(* IEC 61131-3 sources: plc_NativeGateway/tests, 8 files *)

(* ---- NG_TimeResponseTest.st ---- *)
FUNCTION_BLOCK NG_TimeResponseTest
VAR_OUTPUT
    Done : BOOL;
    Passed : UINT;
    FailedChecks : UINT;
    CaseCount : UINT;
END_VAR
VAR
    Parser : NG_JsonParse;
    Reader : NG_TimeResponse;
    Doc : NG_Document;
    Bytes : NG_Bytes;
    CopyString : STRING_TO_BUF;
    Payload : STRING[2048];
    Stage : UINT;
    CaseIndex : UINT := 1;
    Expected : BOOL;
    Retained : BOOL;
    Actual : BOOL;
END_VAR
IF Done THEN RETURN; END_IF;
Parser(Execute:=Stage=1,Length:=TO_UDINT(LEN(Payload)),Buffer:=Bytes,Doc:=Doc);
CASE Stage OF
0:
    CASE CaseIndex OF
        1: Payload:='{"schemaVersion":1,"gatewayId":"PLC-01","requestId":"time-boot-A-1","bootId":"boot-A","sessionId":"session-A","clientMonoMs":10000,"serverReceivedAt":1792739100000,"serverSentAt":1792739100005}'; Expected:=TRUE; Retained:=FALSE;
        2: Payload:='{"schemaVersion":1,"gatewayId":"PLC-01","requestId":"time-boot-A-1","bootId":"boot-A","sessionId":"session-A","clientMonoMs":10000,"serverReceivedAt":1792739100000,"serverSentAt":1792739100005}'; Expected:=TRUE; Retained:=FALSE;
        3: Payload:='{"schemaVersion":1,"gatewayId":"PLC-01","requestId":"time-boot-A-1","bootId":"boot-A","sessionId":"session-A","clientMonoMs":10000,"timestamp":0,"serverReceivedAt":1792739100000,"serverSentAt":1792739100005}'; Expected:=FALSE; Retained:=FALSE;
        4: Payload:='{"schemaVersion":1,"gatewayId":"PLC-01","requestId":"time-boot-A-1","bootId":"boot-A","sessionId":"session-A","clientMonoMs":true,"serverReceivedAt":1792739100000,"serverSentAt":1792739100005}'; Expected:=FALSE; Retained:=FALSE;
        5: Payload:='{"schemaVersion":1,"gatewayId":"PLC-01","requestId":"time-boot-A-1","bootId":"boot-A","sessionId":"session-A","clientMonoMs":10000.0,"serverReceivedAt":1792739100000,"serverSentAt":1792739100005}'; Expected:=FALSE; Retained:=FALSE;
        6: Payload:='{"schemaVersion":1.0,"gatewayId":"PLC-01","requestId":"time-boot-A-1","bootId":"boot-A","sessionId":"session-A","clientMonoMs":10000,"serverReceivedAt":1792739100000,"serverSentAt":1792739100005}'; Expected:=FALSE; Retained:=FALSE;
        7: Payload:='{"schemaVersion":1,"gatewayId":"PLC-01","requestId":"time-boot-A-1","bootId":"boot-A","sessionId":null,"clientMonoMs":10000,"serverReceivedAt":1792739100000,"serverSentAt":1792739100005}'; Expected:=FALSE; Retained:=FALSE;
        8: Payload:='{"schemaVersion":1,"gatewayId":"PLC-01","requestId":"time-boot-A-1","bootId":"boot-A","sessionId":"session-A","clientMonoMs":9007199254740992,"serverReceivedAt":1792739100000,"serverSentAt":1792739100005}'; Expected:=FALSE; Retained:=FALSE;
        9: Payload:='{"schemaVersion":1,"gatewayId":"PLC-01","requestId":"aaaaaaaaaaaaaaaaaaaaaaaaaaaaaaaaaaaaaaaaaaaaaaaaaaaaaaaaaaaaaaaaa","bootId":"boot-A","sessionId":"session-A","clientMonoMs":10000,"serverReceivedAt":1792739100000,"serverSentAt":1792739100005}'; Expected:=FALSE; Retained:=FALSE;
        10: Payload:='{"schemaVersion":1,"gatewayId":"PLC-01","requestId":"a/b","bootId":"boot-A","sessionId":"session-A","clientMonoMs":10000,"serverReceivedAt":1792739100000,"serverSentAt":1792739100005}'; Expected:=FALSE; Retained:=FALSE;
        11: Payload:='{"schemaVersion":1,"gatewayId":"PLC-01","requestId":"time-boot-A-1","bootId":"boot-A","sessionId":"session-A","clientMonoMs":10000,"serverReceivedAt":1792739100000,"serverSentAt":1792739100005}'; Expected:=FALSE; Retained:=TRUE;
        12: Payload:='{"schemaVersion":1,"gatewayId":"other","requestId":"time-boot-A-1","bootId":"boot-A","sessionId":"session-A","clientMonoMs":10000,"serverReceivedAt":1792739100000,"serverSentAt":1792739100005}'; Expected:=FALSE; Retained:=FALSE;
        13: Payload:='{"schemaVersion":1,"gatewayId":"PLC-01","requestId":"time-boot-A-1","bootId":"other","sessionId":"session-A","clientMonoMs":10000,"serverReceivedAt":1792739100000,"serverSentAt":1792739100005}'; Expected:=FALSE; Retained:=FALSE;
        14: Payload:='{"schemaVersion":1,"gatewayId":"PLC-01","requestId":"time-boot-A-1","bootId":"boot-A","sessionId":"other","clientMonoMs":10000,"serverReceivedAt":1792739100000,"serverSentAt":1792739100005}'; Expected:=FALSE; Retained:=FALSE;
        15: Payload:='{"schemaVersion":1,"gatewayId":"PLC-01","requestId":"other","bootId":"boot-A","sessionId":"session-A","clientMonoMs":10000,"serverReceivedAt":1792739100000,"serverSentAt":1792739100005}'; Expected:=FALSE; Retained:=FALSE;
        16: Payload:='{"schemaVersion":1,"gatewayId":"PLC-01","requestId":"time-boot-A-1","bootId":"boot-A","sessionId":"session-A","clientMonoMs":10001,"serverReceivedAt":1792739100000,"serverSentAt":1792739100005}'; Expected:=FALSE; Retained:=FALSE;
        17: Payload:='{"schemaVersion":1,"gatewayId":"PLC-01","requestId":"time-boot-A-1","bootId":"boot-A","sessionId":"session-A","clientMonoMs":10000.0,"serverReceivedAt":1792739100000,"serverSentAt":1792739100005}'; Expected:=FALSE; Retained:=FALSE;
        18: Payload:='{"schemaVersion":1,"gatewayId":"PLC-01","requestId":"time-boot-A-1","bootId":"boot-A","sessionId":"session-A","clientMonoMs":10000,"serverReceivedAt":1792739100000,"serverSentAt":1.0}'; Expected:=FALSE; Retained:=FALSE;
        19: Payload:='{"schemaVersion":1,"gatewayId":"PLC-01","requestId":"time-boot-A-1","bootId":"boot-A","sessionId":"session-A","clientMonoMs":10000,"serverReceivedAt":1792739100000,"serverSentAt":9007199254740992}'; Expected:=FALSE; Retained:=FALSE;
        20: Payload:='{"schemaVersion":1,"gatewayId":"PLC-01","requestId":"time-boot-A-1","bootId":"boot-A","sessionId":"session-A","clientMonoMs":10000,"serverReceivedAt":true,"serverSentAt":1792739100005}'; Expected:=FALSE; Retained:=FALSE;
        21: Payload:='{"schemaVersion":1,"gatewayId":"PLC-01","requestId":"time-boot-A-1","bootId":"boot-A","sessionId":"session-A","clientMonoMs":10000,"serverReceivedAt":1792739100000,"serverSentAt":1792739100005,"timestamp":0}'; Expected:=FALSE; Retained:=FALSE;
        22: Payload:='{"schemaVersion":1,"gatewayId":"PLC-01","requestId":"time-boot-A-1","bootId":"boot-A","sessionId":"session-A","clientMonoMs":10000,"serverReceivedAt":1792739100000,"serverSentAt":1792739100005,"schemaVersion":1}'; Expected:=FALSE; Retained:=FALSE;
        23: Payload:='{"schemaVersion":1e0,"gatewayId":"PLC-01","requestId":"time-boot-A-1","bootId":"boot-A","sessionId":"session-A","clientMonoMs":10000,"serverReceivedAt":1792739100000,"serverSentAt":1792739100005}'; Expected:=FALSE; Retained:=FALSE;
    END_CASE;
    CopyString(REQ:=FALSE,BUF_FORMAT:=FALSE,BUF_OFFS:=0,BUF_CNT:=LEN(Payload),SRC:=Payload,BUFFER:=Bytes);
    CopyString(REQ:=TRUE,BUF_FORMAT:=FALSE,BUF_OFFS:=0,BUF_CNT:=LEN(Payload),SRC:=Payload,BUFFER:=Bytes);
    IF CopyString.DONE THEN Stage:=1; END_IF;
1:
    IF Parser.Error OR Parser.Done THEN
        Actual:=FALSE;
        IF Parser.Done THEN
            Reader(Length:=TO_UDINT(LEN(Payload)),Retained:=Retained,GatewayId:='PLC-01',BootId:='boot-A',
                SessionId:='session-A',RequestId:='time-boot-A-1',ClientMonoMs:=10000,Doc:=Doc,Bytes:=Bytes);
            Actual:=Reader.Valid;
        END_IF;
        IF Actual=Expected THEN Passed:=Passed+1; ELSE FailedChecks:=FailedChecks+1; END_IF;
        CaseCount:=CaseCount+1; Stage:=2;
    END_IF;
2:
    CaseIndex:=CaseIndex+1;
    IF CaseIndex>23 THEN Done:=TRUE; ELSE Stage:=0; END_IF;
END_CASE;
END_FUNCTION_BLOCK

(* ---- audit_facts_test.st ---- *)
PROGRAM Main
VAR
    Buffer : NG_Buffer;
    Event : NG_CaptureEvent;
    AuditRecord : NG_AuditEvent;
    Cursor : NG_SourceCursor;
    Capture : NG_CaptureCore;
    Poll : NG_PollSlot;
    Audit : NG_AuditCapture;
    Decide : NG_AuditDecision;
    Policy : NG_ReportPolicy;
    Checks : ARRAY[1..20] OF BOOL;
    Passed : UINT;
    FailedChecks : UINT;
    Done : BOOL;
    i : UINT;
END_VAR
(* Compile-only harness; no socket, SDK, persistent store, RTC or physical I/O.
   Cold compilation does not execute these assertions. *)
IF Done THEN RETURN; END_IF;
Checks[1]:=SIZEOF(Event)=UDINT#72;
Checks[2]:=SIZEOF(AuditRecord)=UDINT#80;
Checks[3]:=SIZEOF(Cursor)=UDINT#48;
Buffer.AuditEnabled:=TRUE; Buffer.PlatformTime:=TRUE; Buffer.TimeValid:=TRUE;
Event.SampleSeq:=1; Event.ConfigSlot:=1; Event.ConfigGeneration:=1;
Event.CompletedMonoMs:=1000; Event.ClockRevision:=2;
Buffer.DecisionSnapshotMonoMs:=66537; Buffer.ClockRevision:=5;
Audit(Buffer:=Buffer,Event:=Event);
Decide(SampleSeq:=ULINT#1,Decision:=USINT#2,Reason:=USINT#0,ReportSkipped:=ULINT#7,Buffer:=Buffer);
Checks[4]:=Buffer.AuditEvents[1].DecisionFlags=BYTE#63;
Checks[5]:=(Buffer.AuditEvents[1].DecisionDelayLo=1) AND (Buffer.AuditEvents[1].DecisionDelayHi=1);
Checks[6]:=(Buffer.AuditEvents[1].DecisionRevisionDelta=3) AND (Buffer.AuditEvents[1].ReportSkipped=7);
Buffer.DecisionSnapshotMonoMs:=ULINT#16778215; Buffer.ClockRevision:=257;
Audit(Buffer:=Buffer,Event:=Event);
Decide(SampleSeq:=ULINT#1,Decision:=USINT#3,Reason:=USINT#4,ReportSkipped:=ULINT#254,Buffer:=Buffer);
Checks[7]:=(Buffer.AuditEvents[1].DecisionFlags=BYTE#63) AND (Buffer.AuditEvents[1].DecisionDelayLo=65535) AND (Buffer.AuditEvents[1].DecisionDelayHi=255);
Buffer.DecisionSnapshotMonoMs:=ULINT#16778216;
Audit(Buffer:=Buffer,Event:=Event);
Decide(SampleSeq:=ULINT#1,Decision:=USINT#3,Reason:=USINT#4,ReportSkipped:=ULINT#0,Buffer:=Buffer);
Checks[8]:=((Buffer.AuditEvents[1].DecisionFlags AND BYTE#8)=BYTE#0) AND NOT Buffer.AuditFactsComplete;
Buffer.AuditFactsComplete:=TRUE; Buffer.DecisionSnapshotMonoMs:=1000; Buffer.ClockRevision:=258;
Audit(Buffer:=Buffer,Event:=Event);
Decide(SampleSeq:=ULINT#1,Decision:=USINT#3,Reason:=USINT#4,ReportSkipped:=ULINT#255,Buffer:=Buffer);
Checks[9]:=((Buffer.AuditEvents[1].DecisionFlags AND BYTE#16)=BYTE#0) AND ((Buffer.AuditEvents[1].DecisionFlags AND BYTE#32)=BYTE#0);
Buffer.DecisionSnapshotMonoMs:=999; Buffer.ClockRevision:=2;
Audit(Buffer:=Buffer,Event:=Event);
Decide(SampleSeq:=ULINT#1,Decision:=USINT#3,Reason:=USINT#4,ReportSkipped:=ULINT#0,Buffer:=Buffer);
Checks[10]:=(Buffer.AuditEvents[1].DecisionFlags AND BYTE#8)=BYTE#0;
Decide(SampleSeq:=ULINT#1,Decision:=USINT#2,Reason:=USINT#0,ReportSkipped:=ULINT#0,Buffer:=Buffer);
Checks[11]:=NOT Buffer.EvidenceComplete AND (Buffer.AuditEvents[1].Decision=3);
Buffer.EvidenceComplete:=TRUE; Buffer.AuditFactsComplete:=TRUE;
Cursor.NextDueMonoMs:=100;
Poll(NowMs:=ULINT#11100,PeriodMs:=UDINT#5000,Cursor:=Cursor,Buffer:=Buffer);
Checks[12]:=(Poll.NominalDueMs=10100) AND (Cursor.NextDueMonoMs=15100) AND (Cursor.PollSkippedPending=2);
Checks[13]:=Buffer.MissedPollCyclesTotal=2;
Buffer.ActiveSlot:=1; Buffer.LayoutValid:=TRUE; Buffer.NextSampleSeq:=0;
Buffer.SamplingGeneration:=1; Buffer.Configs[1].Generation:=1;
Buffer.Configs[1].Config.Points[1].reportMode:='cyclic';
Buffer.Configs[1].Config.Points[1].reportIntervalMs:=5000;
Buffer.Cursors[1].Enabled:=TRUE; Buffer.Cursors[1].ActivatedMonoMs:=100;
Buffer.Cursors[1].NextDueMonoMs:=15100; Buffer.Cursors[1].PollSkippedPending:=2;
Buffer.ClockRevision:=2; Buffer.TimeValid:=TRUE; Buffer.DecisionSnapshotMonoMs:=11100;
Capture(PointIndex:=UINT#1,Kind:=USINT#1,Quality:=USINT#2,Value:=LREAL#7.0,
    NowMs:=ULINT#11100,NominalDueMs:=ULINT#10100,SystemUtcMs:=ULINT#100000,
    Cursor:=Buffer.Cursors[1],Buffer:=Buffer);
Checks[14]:=(Buffer.AuditEvents[1].Event.PollSkippedBefore=2) AND (Buffer.Cursors[1].PollSkippedPending=0);
Buffer.TimeValid:=FALSE; Buffer.ClockRevision:=3; Buffer.DecisionSnapshotMonoMs:=12000;
Policy(DeferCapacity:=FALSE,Buffer:=Buffer);
Checks[15]:=(Buffer.AuditEvents[1].Decision=3) AND (Buffer.AuditEvents[1].Reason=4);
Checks[16]:=(Buffer.AuditEvents[1].DecisionFlags=BYTE#59) AND (Buffer.AuditEvents[1].DecisionRevisionDelta=1);
Checks[17]:=(Buffer.AuditEvents[1].DecisionDelayLo=900) AND (Buffer.AuditEvents[1].ReportSkipped=2);
Checks[18]:=(Buffer.MissedReportSlotsTotal=2) AND (Buffer.AuditEvents[1].Event.CapturedUtcMs=100000);
Event.SampleSeq:=2; Event.Kind:=2; Event.PointIndex:=1;
Event.CompletedMonoMs:=15200; Event.ClockRevision:=4;
Event.SamplingGeneration:=1; Event.Flags:=WORD#3; Event.Quality:=3;
Buffer.Configs[1].Config.Points[1].pollIntervalMs:=5000;
Buffer.DecisionSnapshotMonoMs:=15210; Buffer.ClockRevision:=4; Buffer.TimeValid:=TRUE;
Buffer.Cursors[1].NextDueMonoMs:=20100;
Audit(Buffer:=Buffer,Event:=Event);
Buffer.Ingress[Buffer.Tail]:=Event; Buffer.Tail:=Buffer.Tail MOD 512+1;
Buffer.IngressCount:=Buffer.IngressCount+1; Buffer.Configs[1].References:=Buffer.Configs[1].References+1;
Policy(DeferCapacity:=FALSE,Buffer:=Buffer);
Checks[19]:=(Buffer.AuditEvents[2].DecisionFlags=BYTE#127) AND (Buffer.AuditEvents[2].ReportSkipped=128);
Event.SampleSeq:=3; Event.CompletedMonoMs:=15300; Event.ClockRevision:=5;
Buffer.ClockRevision:=6; Buffer.TimeValid:=FALSE; Buffer.DecisionSnapshotMonoMs:=15310;
Buffer.Cursors[1].NextDueMonoMs:=655100;
Audit(Buffer:=Buffer,Event:=Event);
Buffer.Ingress[Buffer.Tail]:=Event; Buffer.Tail:=Buffer.Tail MOD 512+1;
Buffer.IngressCount:=Buffer.IngressCount+1; Buffer.Configs[1].References:=Buffer.Configs[1].References+1;
Policy(DeferCapacity:=FALSE,Buffer:=Buffer);
Checks[20]:=((Buffer.AuditEvents[3].DecisionFlags AND BYTE#32)=BYTE#0) AND NOT Buffer.AuditFactsComplete;
FOR i:=1 TO 20 DO
    IF Checks[i] THEN Passed:=Passed+1; ELSE FailedChecks:=FailedChecks+1; END_IF;
END_FOR;
Done:=TRUE;
END_PROGRAM

(* ---- phase1_capture_test.st ---- *)
PROGRAM Main
VAR
    Buffer : NG_Buffer;
    Samples : ARRAY[1..320] OF NG_Sample;
    Config : NG_Config;
    Selector : NG_ConfigSlot;
    Source : NG_SourceState;
    Result : NG_SourceResult;
    Poll : NG_PollSlot;
    Capture : NG_Capture;
    Compare : NG_SameConfig;
    Stage : INT;
    Passed : UDINT;
    FailedChecks : UDINT;
    Done : BOOL;
    Check : BOOL;
    Checks : ARRAY[1..40] OF BOOL;
    RecordBytes : UDINT;
    BufferBytes : UDINT;
    BudgetBytes : UDINT;
    DummyPacket : NG_Packet;
    Packets : ARRAY[1..16] OF NG_Packet;
    Values : NG_Json;
    TxPayload : NG_Json;
    Item : STRING[1024];
    Point : NG_Point;
    Sample : NG_Sample;
    Tx : NG_Bytes;
    Rx : NG_Bytes;
    n : INT;
    PreviousSeq : ULINT;
    PreviousCaptured : ULINT;
    OldSlot : UINT;
    OldGeneration : UDINT;
    HashBefore : ULINT;
END_VAR
IF Done THEN RETURN; END_IF;
Check:=FALSE;
CASE Stage OF
0:
    RecordBytes:=SIZEOF(Buffer.Scratch); BufferBytes:=SIZEOF(Buffer);
    BudgetBytes:=BufferBytes+SIZEOF(Packets)+SIZEOF(Samples)+SIZEOF(Values)+SIZEOF(Item)+SIZEOF(TxPayload)+SIZEOF(DummyPacket)+SIZEOF(Sample)+SIZEOF(Point)+SIZEOF(Tx)+SIZEOF(Rx)+UDINT#16384+UDINT#135680+UDINT#65536;
    Buffer.LayoutValid:=BudgetBytes<=UDINT#4194304;
    Config.Version:=1; Config.MessageId:='capture-test-1'; Config.enabled:=TRUE;
    Config.DeviceCount:=1; Config.PointCount:=3;
    Config.Devices[1].deviceId:='D1'; Config.Devices[1].PointStart:=1; Config.Devices[1].PointCount:=3;
    FOR n:=1 TO 3 DO Config.Points[n].enabled:=TRUE; Config.Points[n].pollIntervalMs:=1000; END_FOR;
    Config.Points[1].pointId:='P1'; Config.Points[2].pointId:='P2'; Config.Points[3].pointId:='P3';
    Selector(GatewayId:='TEST',CaptureBootId:='BOOT',Config:=Config,Buffer:=Buffer);
    Buffer.ActiveSlot:=Selector.Slot; Buffer.Configs[Selector.Slot].Reserved:=FALSE; Buffer.SamplingGeneration:=1;
    Check:=(Selector.Slot>0) AND Buffer.LayoutValid;
1: (* UNKNOWN once; nominal slot is absent; O comes from activation. *)
    Source(Index:=1,Enabled:=TRUE,NowMs:=100,UnixMs:=100000,StaleAfterMs:=3000,CheckStale:=FALSE,Samples:=Samples,Buffer:=Buffer);
    Check:=Source.Accepted AND (Buffer.IngressCount=1) AND (Buffer.Ingress[1].Kind=2) AND (Buffer.Ingress[1].Quality=1) AND (Buffer.Cursors[1].NextDueMonoMs=100) AND ((Buffer.Ingress[1].Flags AND WORD#4)=WORD#0);
2:
    Source(Index:=1,Enabled:=TRUE,NowMs:=200,UnixMs:=100000,StaleAfterMs:=3000,CheckStale:=TRUE,Samples:=Samples,Buffer:=Buffer);
    Check:=(Buffer.CapturedEventsTotal=1) AND (Buffer.Cursors[1].NextDueMonoMs=100);
3: (* Final BAD counts as physical liveness. *)
    Poll(NowMs:=1100,PeriodMs:=1000,Cursor:=Buffer.Cursors[1],Buffer:=Buffer);
    Result(Index:=1,Value:=LREAL#123.0,Quality:='BAD_TIMEOUT',NowMs:=1110,UnixMs:=101000,NominalDueMs:=Poll.NominalDueMs,ConfigSlot:=Buffer.ActiveSlot,ConfigGeneration:=Buffer.Configs[Buffer.ActiveSlot].Generation,SamplingGeneration:=1,Samples:=Samples,Buffer:=Buffer);
    Check:=Result.Accepted AND (Buffer.MissedPollCyclesTotal=1) AND (Buffer.Ingress[2].Value=0) AND (Buffer.Ingress[2].NominalDueMonoMs=1100) AND (Buffer.Cursors[1].NextDueMonoMs=2100);
4:
    Source(Index:=1,Enabled:=TRUE,NowMs:=4000,UnixMs:=101000,StaleAfterMs:=3000,CheckStale:=TRUE,Samples:=Samples,Buffer:=Buffer);
    Check:=(Buffer.CapturedEventsTotal=2) AND (Samples[1].Quality='BAD_TIMEOUT');
5:
    Result(Index:=1,Value:=LREAL#0.0,Quality:='BAD_TIMEOUT',NowMs:=4100,UnixMs:=101000,NominalDueMs:=2100,ConfigSlot:=Buffer.ActiveSlot,ConfigGeneration:=Buffer.Configs[Buffer.ActiveSlot].Generation,SamplingGeneration:=1,Samples:=Samples,Buffer:=Buffer);
    Source(Index:=1,Enabled:=TRUE,NowMs:=4100,UnixMs:=101000,StaleAfterMs:=3000,CheckStale:=TRUE,Samples:=Samples,Buffer:=Buffer);
    Check:=(Buffer.CapturedEventsTotal=3) AND (Buffer.SourceTimestampRepeatTotal=1) AND (Samples[1].Quality='BAD_TIMEOUT');
6: (* STALE at the exact boundary, once. *)
    Source(Index:=1,Enabled:=TRUE,NowMs:=7100,UnixMs:=107000,StaleAfterMs:=3000,CheckStale:=TRUE,Samples:=Samples,Buffer:=Buffer);
    Check:=(Buffer.CapturedEventsTotal=4) AND (Buffer.Ingress[4].Kind=2) AND (Buffer.Ingress[4].Quality=3) AND (Buffer.Ingress[4].CompletedMonoMs=7100);
7:
    Source(Index:=1,Enabled:=TRUE,NowMs:=7200,UnixMs:=108000,StaleAfterMs:=3000,CheckStale:=TRUE,Samples:=Samples,Buffer:=Buffer);
    Check:=(Buffer.CapturedEventsTotal=4);
8: (* GOOD scalar is frozen, never rescaled by capture. *)
    Result(Index:=1,Value:=LREAL#42.25,Quality:='GOOD',NowMs:=7300,UnixMs:=109000,NominalDueMs:=3100,ConfigSlot:=Buffer.ActiveSlot,ConfigGeneration:=Buffer.Configs[Buffer.ActiveSlot].Generation,SamplingGeneration:=1,Samples:=Samples,Buffer:=Buffer);
    Check:=(Buffer.CapturedEventsTotal=5) AND (Buffer.Ingress[5].Value=LREAL#42.25) AND (Buffer.Ingress[5].CapturedUtcMs=109000) AND ((Buffer.Ingress[5].Flags AND WORD#10)=WORD#8);
9: (* Equal RTC remains two events. *)
    Result(Index:=1,Value:=LREAL#43.25,Quality:='GOOD',NowMs:=7310,UnixMs:=109000,NominalDueMs:=4100,ConfigSlot:=Buffer.ActiveSlot,ConfigGeneration:=Buffer.Configs[Buffer.ActiveSlot].Generation,SamplingGeneration:=1,Samples:=Samples,Buffer:=Buffer);
    Check:=(Buffer.CapturedEventsTotal=6) AND (Buffer.SourceTimestampRepeatTotal=2) AND (Buffer.Ingress[5].Value=LREAL#42.25) AND (Buffer.Ingress[6].Value=LREAL#43.25);
10: (* RTC invalid is null, no later backfill. *)
    Result(Index:=1,Value:=LREAL#44.0,Quality:='GOOD',NowMs:=7400,UnixMs:=0,NominalDueMs:=5100,ConfigSlot:=Buffer.ActiveSlot,ConfigGeneration:=Buffer.Configs[Buffer.ActiveSlot].Generation,SamplingGeneration:=1,Samples:=Samples,Buffer:=Buffer);
    Check:=((Buffer.Ingress[7].Flags AND WORD#1)=WORD#0) AND (Buffer.Ingress[7].CapturedUtcMs=0) AND (Buffer.Ingress[5].CapturedUtcMs=109000);
11: (* Per-point missed slots in an N-point logical block. *)
    FOR n:=2 TO 3 DO
        Source(Index:=TO_UINT(n),Enabled:=TRUE,NowMs:=100,UnixMs:=100000,StaleAfterMs:=3000,CheckStale:=FALSE,Samples:=Samples,Buffer:=Buffer);
        Poll(NowMs:=3100,PeriodMs:=1000,Cursor:=Buffer.Cursors[n],Buffer:=Buffer);
    END_FOR;
    Check:=(Buffer.MissedPollCyclesTotal=7) AND (Buffer.Cursors[2].NextDueMonoMs=4100) AND (Buffer.Cursors[3].NextDueMonoMs=4100);
12: (* Old read revoked, no new event or source-view mutation. *)
    PreviousCaptured:=Buffer.CapturedEventsTotal;
    Result(Index:=1,Value:=LREAL#99.0,Quality:='GOOD',NowMs:=7500,UnixMs:=110000,NominalDueMs:=6100,ConfigSlot:=Buffer.ActiveSlot,ConfigGeneration:=0,SamplingGeneration:=1,Samples:=Samples,Buffer:=Buffer);
    Check:=NOT Result.Accepted AND (Buffer.CapturedEventsTotal=PreviousCaptured) AND (Samples[1].Value=LREAL#44.0) AND (Buffer.CancelledReadsTotal=1) AND (Buffer.CancellationReason=2);
13: (* Idempotent config application keeps slot and sampling origin. *)
    OldSlot:=Buffer.ActiveSlot; OldGeneration:=Buffer.Configs[OldSlot].Generation;
    Selector(GatewayId:='TEST',CaptureBootId:='BOOT',Config:=Config,Buffer:=Buffer);
    Check:=(Selector.Slot=OldSlot) AND (Buffer.Configs[OldSlot].Generation=OldGeneration) AND (Buffer.Configs[OldSlot].References=Buffer.IngressCount);
14: (* All versions retained, old slot is immutable. *)
    Config.Version:=2; Config.MessageId:='capture-test-2'; Config.Points[1].scale:=2;
    Selector(GatewayId:='TEST',CaptureBootId:='BOOT',Config:=Config,Buffer:=Buffer);
    Buffer.ActiveSlot:=Selector.Slot; Buffer.Configs[Selector.Slot].Reserved:=FALSE; Buffer.SamplingGeneration:=2;
    Check:=(Selector.Slot<>OldSlot) AND (Buffer.Configs[OldSlot].Config.Version=1) AND (Buffer.Ingress[5].ConfigGeneration=OldGeneration) AND (Buffer.Ingress[5].Value=LREAL#42.25);
15:
    Source(Index:=1,Enabled:=TRUE,NowMs:=8000,UnixMs:=111000,StaleAfterMs:=3000,CheckStale:=FALSE,Samples:=Samples,Buffer:=Buffer);
    Check:=Source.Accepted AND (Buffer.Cursors[1].NextDueMonoMs=8000) AND (Samples[1].Quality='UNKNOWN');
16: (* Pin all four dictionaries. Fifth version cannot replace current/history. *)
    FOR n:=3 TO 4 DO
        Config.Version:=TO_ULINT(n);
        Selector(GatewayId:='TEST',CaptureBootId:='BOOT',Config:=Config,Buffer:=Buffer);
        Buffer.ActiveSlot:=Selector.Slot; Buffer.Configs[Selector.Slot].Reserved:=FALSE;
        Buffer.SamplingGeneration:=TO_ULINT(n);
        Capture(PointIndex:=1,Kind:=2,Quality:=1,Value:=LREAL#0.0,NowMs:=9000,NominalDueMs:=0,SystemUtcMs:=112000,Buffer:=Buffer);
    END_FOR;
    OldSlot:=Buffer.ActiveSlot; Config.Version:=5;
    Selector(GatewayId:='TEST',CaptureBootId:='BOOT',Config:=Config,Buffer:=Buffer);
    Check:=(Selector.Slot=0) AND (Buffer.ActiveSlot=OldSlot) AND (Buffer.Configs[OldSlot].Config.Version=4) AND (Buffer.Configs[1].Config.Version=1);
17: (* Queue fill one bounded capture per scan. *)
    IF Buffer.IngressCount<512 THEN
        Capture(PointIndex:=1,Kind:=1,Quality:=2,Value:=LREAL#12.0,NowMs:=10000,NominalDueMs:=10000,SystemUtcMs:=112000,Buffer:=Buffer);
        RETURN;
    END_IF;
    PreviousSeq:=Buffer.NextSampleSeq; PreviousCaptured:=Buffer.CapturedEventsTotal;
    Check:=(Buffer.CaptureOverflowEventsTotal=0);
18:
    Capture(PointIndex:=1,Kind:=1,Quality:=2,Value:=LREAL#99.0,NowMs:=10001,NominalDueMs:=10000,SystemUtcMs:=112000,Buffer:=Buffer);
    Check:=NOT Capture.Accepted AND (Buffer.IngressCount=512) AND (Buffer.CaptureOverflowEventsTotal=1) AND (Buffer.UndecidedLostEventsTotal=1) AND (Buffer.NextSampleSeq=PreviousSeq+1) AND (Buffer.CapturedEventsTotal=PreviousCaptured+1) AND (Buffer.Ingress[5].Value=LREAL#42.25) AND (Buffer.Gaps[1].PointId='P1');
19: (* Bounded detail ring; totals remain exact. *)
    FOR n:=1 TO 64 DO
        Capture(PointIndex:=1,Kind:=1,Quality:=5,Value:=LREAL#0.0,NowMs:=10002,NominalDueMs:=10000,SystemUtcMs:=112000,Buffer:=Buffer);
    END_FOR;
    Check:=(Buffer.CaptureOverflowEventsTotal=65) AND (Buffer.UndecidedLostEventsTotal=65) AND Buffer.DetailTruncated AND (Buffer.GapIndex=1);
20:
    Check:=(NG_SafeAdd(ULINT#9007199254740990,ULINT#10)=ULINT#9007199254740991) AND (NG_SafeAdd(ULINT#7,ULINT#4)=11);
21: (* Exhausted sample identity fails closed, never wraps. *)
    Buffer.NextSampleSeq:=ULINT#9007199254740991; PreviousCaptured:=Buffer.CapturedEventsTotal;
    Capture(PointIndex:=1,Kind:=1,Quality:=2,Value:=LREAL#99.0,NowMs:=11000,NominalDueMs:=11000,SystemUtcMs:=113000,Buffer:=Buffer);
    Check:=NOT Capture.Accepted AND Buffer.CaptureStopped AND (Buffer.CapturedEventsTotal=PreviousCaptured) AND (Buffer.NextSampleSeq=ULINT#9007199254740991);
ELSE Done:=TRUE; RETURN;
END_CASE;
Checks[Stage+1]:=Check;
IF Check THEN Passed:=Passed+1; ELSE FailedChecks:=FailedChecks+1; END_IF;
Stage:=Stage+1;
END_PROGRAM

(* ---- phase1_diagnostics_test.st ---- *)
PROGRAM Main
VAR
    Buffer : NG_Buffer;
    Capture : NG_Capture;
    Policy : NG_ReportPolicy;
    Drain : NG_AuditDrain;
    Associate : NG_AuditAssociation;
    Diagnostics : NG_Diagnostics;
    Stage : INT;
    Checks : ARRAY[1..16] OF BOOL;
    Passed : UINT;
    FailedChecks : UINT;
    Done : BOOL;
    i : INT;
END_VAR
IF Done THEN RETURN; END_IF;
CASE Stage OF
0:
    Buffer.ActiveSlot:=1; Buffer.LayoutValid:=TRUE; Buffer.SamplingGeneration:=1;
    Buffer.Configs[1].Generation:=1; Buffer.Configs[1].GatewayId:='test-gw'; Buffer.Configs[1].CaptureBootId:='test-boot';
    Buffer.Configs[1].Config.Version:=13; Buffer.Configs[1].Config.DeviceCount:=1;
    Buffer.Configs[1].Config.PointCount:=1; Buffer.Configs[1].Config.Devices[1].deviceId:='device';
    Buffer.Configs[1].Config.Devices[1].PointStart:=1; Buffer.Configs[1].Config.Devices[1].PointCount:=1;
    Buffer.Configs[1].Config.Points[1].pointId:='point'; Buffer.Configs[1].Config.Points[1].reportMode:='cyclic';
    Buffer.Configs[1].Config.Points[1].reportIntervalMs:=5000; Buffer.Cursors[1].Enabled:=TRUE;
    Buffer.AuditEnabled:=TRUE; Buffer.LayoutBytes:=SIZEOF(Buffer); Buffer.RecordBytes:=SIZEOF(Buffer.Scratch);
    Diagnostics(BootId:='test-boot',GatewayId:='test-gw',NowMs:=ULINT#1000,Force:=TRUE,Buffer:=Buffer);
    Checks[1]:=Buffer.Diagnostics.RestartLossUnknown AND NOT Buffer.Diagnostics.AccountingComplete AND (Buffer.Diagnostics.Totals[16]=1) AND NOT Buffer.Diagnostics.LastGapCountKnown;
    Checks[2]:=NOT Buffer.Diagnostics.HasPendingAge AND (Buffer.Diagnostics.PendingEvents=0) AND (Buffer.Diagnostics.Revision MOD 2=0);
    Capture(PointIndex:=UINT#1,Kind:=USINT#1,Quality:=USINT#2,Value:=LREAL#12.5,NowMs:=ULINT#10,NominalDueMs:=ULINT#0,SystemUtcMs:=ULINT#1000,Buffer:=Buffer);
    Checks[3]:=(Buffer.AuditWriteSeq=1) AND (Buffer.AuditEvents[1].Event.Value=LREAL#12.5) AND (Buffer.AuditEvents[1].Decision=0) AND (Buffer.Configs[1].References=2);
    Buffer.AuditAckBootId:='test-boot'; Buffer.AuditAckSeq:=1; Drain(BootId:='test-boot',Buffer:=Buffer);
    Checks[4]:=(Buffer.AuditReadSeq=0) AND (Buffer.Configs[1].References=2);
    Policy(Buffer:=Buffer);
    Checks[5]:=(Buffer.AuditEvents[1].Decision=2) AND (Buffer.OwnedCount=1) AND (Buffer.Configs[1].References=2);
    Buffer.AuditAckBootId:='old-boot'; Drain(BootId:='test-boot',Buffer:=Buffer);
    Checks[6]:=(Buffer.AuditReadSeq=0) AND (Buffer.Configs[1].References=2);
    Buffer.AuditAckBootId:='test-boot'; Drain(BootId:='test-boot',Buffer:=Buffer);
    Checks[7]:=(Buffer.AuditReadSeq=1) AND (Buffer.Configs[1].References=1) AND (Buffer.OwnedCount=1);
    Drain(BootId:='test-boot',Buffer:=Buffer);
    Checks[8]:=(Buffer.Configs[1].References=1);
    Buffer.BatchOwners[1].ConfigSlot:=1; Buffer.BatchOwners[1].Count:=1;
    Buffer.BatchOwners[1].Category:=2; Buffer.BatchOwners[1].Digest:='frozen-hash';
    Buffer.BatchRefs[1]:=1; Buffer.BatchGenerations[1]:=7;
    Associate(Slot:=UINT#1,MessageId:='frozen-message',Buffer:=Buffer);
    Checks[9]:=(Buffer.AssociationWriteSeq=1) AND (Buffer.Associations[1].SampleSeqs[1]=1) AND (Buffer.Associations[1].BatchGeneration=7) AND (Buffer.Configs[1].References=2);
    Buffer.BatchRefs[1]:=0; Buffer.BatchOwners[1].Digest:='changed';
    Checks[10]:=(Buffer.Associations[1].SampleSeqs[1]=1) AND (Buffer.Associations[1].Digest='frozen-hash');
    Buffer.AssociationAckBootId:='test-boot'; Buffer.AssociationAckSeq:=1; Drain(BootId:='test-boot',Buffer:=Buffer);
    Checks[11]:=(Buffer.AssociationReadSeq=1) AND (Buffer.Configs[1].References=1);
    Stage:=1;
1:
    (* Fill the evidence ring independently of business owners. The following
       cyclic events are filtered: only the audit ring remains pinned. *)
    FOR i:=1 TO 64 DO
        Capture(PointIndex:=UINT#1,Kind:=USINT#1,Quality:=USINT#2,Value:=LREAL#12.5,NowMs:=ULINT#100,NominalDueMs:=ULINT#0,SystemUtcMs:=ULINT#1100,Buffer:=Buffer);
    END_FOR;
    Policy(Buffer:=Buffer);
    IF Buffer.AuditWriteSeq>=513 THEN Stage:=2; END_IF;
2:
    Capture(PointIndex:=UINT#1,Kind:=USINT#1,Quality:=USINT#2,Value:=LREAL#12.5,NowMs:=ULINT#100,NominalDueMs:=ULINT#0,SystemUtcMs:=ULINT#1100,Buffer:=Buffer);
    Policy(Buffer:=Buffer);
    Checks[12]:=(Buffer.AuditDropped=1) AND NOT Buffer.EvidenceComplete AND (Buffer.OwnedCount=1) AND (Buffer.KnownUnsentEventsTotal=0) AND (Buffer.UndecidedLostEventsTotal=0);
    Checks[13]:=(Buffer.AuditReadSeq=2) AND (Buffer.Configs[1].References=513) AND (Buffer.AuditEvents[2].Event.SampleSeq=514);
    Diagnostics(BootId:='test-boot',GatewayId:='test-gw',NowMs:=ULINT#2000,Force:=TRUE,Buffer:=Buffer);
    Checks[14]:=(Buffer.Diagnostics.Totals[1]=514) AND (Buffer.Diagnostics.Totals[2]=1) AND (Buffer.Diagnostics.Totals[3]=513) AND (Buffer.Diagnostics.AuditDropped=1) AND (Buffer.Diagnostics.PendingEvents=1);
    Buffer.IngressCount:=2; Buffer.DeadRetainedEvents:=1; Buffer.OwnedCount:=3; Buffer.UncertainRetainedEvents:=1;
    Diagnostics(BootId:='test-boot',GatewayId:='test-gw',NowMs:=ULINT#3000,Force:=TRUE,Buffer:=Buffer);
    Checks[15]:=(Buffer.Diagnostics.PendingEvents=3) AND (Buffer.Diagnostics.DeadEvents=1) AND (Buffer.Diagnostics.UncertainRetainedEvents=1);
    Checks[16]:=(Buffer.Diagnostics.Revision MOD 2=0) AND (Buffer.Diagnostics.AllocatedBytes=SIZEOF(Buffer)) AND (Buffer.Diagnostics.MaxBytes=4194304);
    FOR i:=1 TO 16 DO IF Checks[i] THEN Passed:=Passed+1; ELSE FailedChecks:=FailedChecks+1; END_IF; END_FOR;
    Done:=TRUE;
END_CASE;
END_PROGRAM

(* ---- phase1_performance_test.st ---- *)
PROGRAM Main
VAR_EXTERNAL
    ESM_DATA : ESM_DAT;
END_VAR
VAR
    Buffer : NG_Buffer;
    Samples : ARRAY[1..320] OF NG_Sample;
    Packets : ARRAY[1..16] OF NG_Packet;
    State : NG_SourceState;
    Result : NG_SourceResult;
    Policy : NG_ReportPolicy;
    Maintenance : NG_BufferMaintenance;
    Builder : NG_BatchBuilder;
    Delivery : NG_DeliveryParallel;
    Drain : NG_AuditDrain;
    Diagnostics : NG_Diagnostics;
    Sequence : ULINT;
    Tick : ULINT;
    Scan : UDINT;
    Stage : UINT;
    SamplesMeasured : UDINT;
    SetupUs : LINT;
    SourceStartupUs : LINT;
    LastUs : LINT;
    MaxUs : LINT;
    MinUs : LINT := LINT#9223372036854775807;
    SumUs : ULINT;
    OverOneMs : UDINT;
    OverPeriod : UDINT;
    Done : BOOL;
    d : INT;
    p : INT;
    slot : UINT;
    SubmitAck : BOOL;
    AckId : NG_Id;
    AckQueue : ARRAY[1..8] OF NG_Id;
    AckHead : UINT := 1;
    AckTail : UINT := 1;
    AckCount : UINT;
    ProfileStart : ULINT;
    ProfileWhole : ULINT;
    ProfileDelta : ULINT;
    ProfileMax : ARRAY[1..8] OF ULINT;
    ProfileSum : ARRAY[1..8] OF ULINT;
    ProfileLast : ARRAY[1..8] OF ULINT;
    ProfileIndex : INT;
END_VAR
IF Done THEN RETURN; END_IF;
IF Stage=0 THEN
    Buffer.ActiveSlot:=1; Buffer.SamplingGeneration:=1; Buffer.LayoutValid:=TRUE; Buffer.AuditEnabled:=TRUE;
    Buffer.Configs[1].Generation:=1; Buffer.Configs[1].GatewayId:='test-gw'; Buffer.Configs[1].CaptureBootId:='test-boot';
    Buffer.Configs[1].Config.Version:=13; Buffer.Configs[1].Config.DeviceCount:=50; Buffer.Configs[1].Config.PointCount:=250;
    Buffer.Configs[1].Config.enabled:=TRUE; Buffer.Configs[1].Config.maxBatchPoints:=64;
    Buffer.RecordBytes:=SIZEOF(Buffer.Scratch); Buffer.LayoutBytes:=SIZEOF(Buffer);
    FOR d:=1 TO 50 DO
        Buffer.Configs[1].Config.Devices[d].deviceId:=CONCAT('d-2113457017974222',TO_STRING(850+d,'{0:d}'));
        Buffer.Configs[1].Config.Devices[d].enabled:=TRUE;
        Buffer.Configs[1].Config.Devices[d].PointStart:=(d-1)*5+1; Buffer.Configs[1].Config.Devices[d].PointCount:=5;
    END_FOR;
    FOR p:=1 TO 250 DO
        Buffer.Configs[1].Config.Points[p].pointId:=CONCAT('p-2113457019169599',TO_STRING(490+p,'{0:d}'));
        Buffer.Configs[1].Config.Points[p].enabled:=TRUE;
        Buffer.Configs[1].Config.Points[p].reportMode:='cyclic'; Buffer.Configs[1].Config.Points[p].reportIntervalMs:=5000;
        Buffer.Configs[1].Config.Points[p].dataType:='float32';
    END_FOR;
    Stage:=1; RETURN;
END_IF;
Scan:=Scan+1; Tick:=TO_ULINT(Scan-1)*20;
LastUs:=ESM_DATA.ESM_INFOS[1].TASK_INFOS[1].LAST_EXEC_DURATION;
IF Scan=1 THEN SetupUs:=LastUs;
ELSE
    IF Scan=2 THEN SourceStartupUs:=LastUs; END_IF;
    SamplesMeasured:=SamplesMeasured+1; MaxUs:=MAX(MaxUs,LastUs); MinUs:=MIN(MinUs,LastUs); SumUs:=SumUs+TO_ULINT(LastUs);
    IF LastUs>1000 THEN OverOneMs:=OverOneMs+1; END_IF;
    IF LastUs>20000 THEN OverPeriod:=OverPeriod+1; END_IF;
END_IF;
ProfileWhole:=GET_MICROSECONDS(TRUE); ProfileStart:=ProfileWhole; Buffer.WorkDeadlineUs:=ProfileWhole+ULINT#850;
Drain(BootId:='test-boot',Buffer:=Buffer);
FOR p:=1 TO 250 DO
IF (Buffer.Cursors[p].Generation<>Buffer.SamplingGeneration) OR NOT Buffer.Cursors[p].Enabled OR
   ((Buffer.Cursors[p].Quality<>3) AND (Tick>=Buffer.Cursors[p].LastPhysicalMonoMs+ULINT#30000)) THEN State(Index:=TO_UINT(p),Enabled:=TRUE,NowMs:=Tick,UnixMs:=ULINT#1792840000000+Tick,StaleAfterMs:=UDINT#30000,CheckStale:=TRUE,Samples:=Samples,Buffer:=Buffer); END_IF; END_FOR;
ProfileLast[1]:=GET_MICROSECONDS(TRUE)-ProfileStart; ProfileStart:=GET_MICROSECONDS(TRUE);
(* 50 parallel device completions on five scans per 5 seconds: 250/5s.
   This fixture has no sockets/SDK/MQTT. Its ACKs test logic cost only. *)
IF (Scan>=11) AND ((Scan-11) MOD 250<5) THEN
    FOR d:=1 TO 50 DO
        p:=(d-1)*5+TO_INT((Scan-11) MOD 250)+1;
        Result(Index:=TO_UINT(p),Value:=LREAL#123.125,Quality:='GOOD',NowMs:=Tick,UnixMs:=ULINT#1792840000000+Tick,
            NominalDueMs:=Tick-Tick MOD 5000,ConfigSlot:=UINT#1,ConfigGeneration:=UDINT#1,SamplingGeneration:=ULINT#1,Samples:=Samples,Buffer:=Buffer);
    END_FOR;
END_IF;
ProfileLast[2]:=GET_MICROSECONDS(TRUE)-ProfileStart; ProfileStart:=GET_MICROSECONDS(TRUE);
Maintenance(GateOpen:=TRUE,NowMs:=Tick,Buffer:=Buffer,Packets:=Packets);
ProfileLast[3]:=GET_MICROSECONDS(TRUE)-ProfileStart; ProfileStart:=GET_MICROSECONDS(TRUE);
Policy(Buffer:=Buffer);
ProfileLast[4]:=GET_MICROSECONDS(TRUE)-ProfileStart; ProfileStart:=GET_MICROSECONDS(TRUE);
IF Scan MOD 2=0 THEN
Builder(GateOpen:=TRUE,NowMs:=Tick,UnixMs:=ULINT#1792840000000+Tick,GatewayId:='test-gw',BootId:='test-boot',BatchIntervalMs:=UDINT#1000,Buffer:=Buffer,Packets:=Packets,Sequence:=Sequence);
ProfileLast[5]:=GET_MICROSECONDS(TRUE)-ProfileStart; ProfileStart:=GET_MICROSECONDS(TRUE);
SubmitAck:=FALSE; AckId:='';
IF (AckCount>0) AND NOT Delivery.AckBusy THEN
    SubmitAck:=TRUE; AckId:=AckQueue[AckHead]; AckHead:=AckHead MOD 8+1; AckCount:=AckCount-1;
END_IF;
Delivery(GateOpen:=TRUE,NowMs:=Tick,GatewayId:='test-gw',BootId:='test-boot',SubmitAck:=SubmitAck,AckMessageId:=AckId,
    AckStored:=TRUE,AckRetryable:=FALSE,AckCodes:='',Buffer:=Buffer,Packets:=Packets);
slot:=Delivery.SendSlot;
IF slot>0 THEN
    IF (Tick>=Buffer.NextSendAt) AND (Tick>=Packets[slot].RetryAtMs) THEN
        Packets[slot].WasSent:=TRUE; Packets[slot].RetryAtMs:=Tick+30000; Buffer.NextSendAt:=Tick+334;
        Buffer.PreferSend:=USINT#3-Buffer.BatchOwners[slot].Category;
        IF AckCount>=8 THEN Buffer.CaptureStopped:=TRUE;
        ELSE AckQueue[AckTail]:=Packets[slot].MessageId; AckTail:=AckTail MOD 8+1; AckCount:=AckCount+1; END_IF;
    END_IF;
END_IF;
ProfileLast[6]:=GET_MICROSECONDS(TRUE)-ProfileStart; ProfileStart:=GET_MICROSECONDS(TRUE);
ELSE
SubmitAck:=FALSE; AckId:='';
IF (AckCount>0) AND NOT Delivery.AckBusy THEN
    SubmitAck:=TRUE; AckId:=AckQueue[AckHead]; AckHead:=AckHead MOD 8+1; AckCount:=AckCount-1;
END_IF;
Delivery(GateOpen:=TRUE,NowMs:=Tick,GatewayId:='test-gw',BootId:='test-boot',SubmitAck:=SubmitAck,AckMessageId:=AckId,
    AckStored:=TRUE,AckRetryable:=FALSE,AckCodes:='',Buffer:=Buffer,Packets:=Packets);
slot:=Delivery.SendSlot;
IF slot>0 THEN
    IF (Tick>=Buffer.NextSendAt) AND (Tick>=Packets[slot].RetryAtMs) THEN
        Packets[slot].WasSent:=TRUE; Packets[slot].RetryAtMs:=Tick+30000; Buffer.NextSendAt:=Tick+334;
        Buffer.PreferSend:=USINT#3-Buffer.BatchOwners[slot].Category;
        IF AckCount>=8 THEN Buffer.CaptureStopped:=TRUE;
        ELSE AckQueue[AckTail]:=Packets[slot].MessageId; AckTail:=AckTail MOD 8+1; AckCount:=AckCount+1; END_IF;
    END_IF;
END_IF;
ProfileLast[6]:=GET_MICROSECONDS(TRUE)-ProfileStart; ProfileStart:=GET_MICROSECONDS(TRUE);
Builder(GateOpen:=TRUE,NowMs:=Tick,UnixMs:=ULINT#1792840000000+Tick,GatewayId:='test-gw',BootId:='test-boot',BatchIntervalMs:=UDINT#1000,Buffer:=Buffer,Packets:=Packets,Sequence:=Sequence);
ProfileLast[5]:=GET_MICROSECONDS(TRUE)-ProfileStart; ProfileStart:=GET_MICROSECONDS(TRUE);
END_IF;
Diagnostics(BootId:='test-boot',GatewayId:='test-gw',NowMs:=Tick,Force:=FALSE,Buffer:=Buffer);
Buffer.AuditAckBootId:='test-boot'; Buffer.AuditAckSeq:=Buffer.AuditWriteSeq;
Buffer.AssociationAckBootId:='test-boot'; Buffer.AssociationAckSeq:=Buffer.AssociationWriteSeq;
ProfileLast[7]:=GET_MICROSECONDS(TRUE)-ProfileStart;
ProfileLast[8]:=GET_MICROSECONDS(TRUE)-ProfileWhole;
FOR ProfileIndex:=1 TO 8 DO
    ProfileMax[ProfileIndex]:=MAX(ProfileMax[ProfileIndex],ProfileLast[ProfileIndex]);
    ProfileSum[ProfileIndex]:=ProfileSum[ProfileIndex]+ProfileLast[ProfileIndex];
END_FOR;
IF SamplesMeasured>=600 THEN Done:=TRUE; END_IF;
END_PROGRAM

(* ---- phase1_pipeline_slice_checks.st ---- *)
(* Included only by --slice-assertions in the no-I/O harness. *)
110:
    EndBatch(Slot:=UINT#1,Outcome:=USINT#2,Reason:=USINT#0,NowMs:=Tick,Buffer:=Buffer,Packets:=Packets);
    Capture(PointIndex:=UINT#2,Kind:=USINT#1,Quality:=USINT#2,Value:=LREAL#1.0,NowMs:=ULINT#15010,NominalDueMs:=ULINT#15000,SystemUtcMs:=ULINT#16000,Buffer:=Buffer);
    Policy(Buffer:=Buffer); phaseTicks:=0; Stage:=111;
111:
    Buffer.WorkDeadlineUs:=0;
    Builder(SliceTestHold:=TRUE,GateOpen:=TRUE,NowMs:=Tick,UnixMs:=ULINT#17000,GatewayId:='test-gw',BootId:='test-boot',BatchIntervalMs:=UDINT#1,Buffer:=Buffer,Packets:=Packets,Sequence:=Sequence);
    phaseTicks:=phaseTicks+1;
    IF Builder.SliceTestPending OR (phaseTicks>500) THEN
        savedGeneration:=Buffer.RecordGenerations[Buffer.QueueHead[2]]; firstSlot:=Buffer.QueueHead[2];
        CheckIndex:=47; Check:=Builder.SliceTestPending AND (Buffer.BatchOwners[1].Count=0) AND (firstSlot>0) AND (Buffer.RecordStates[firstSlot]=1);
        Maintenance(GateOpen:=FALSE,NowMs:=ULINT#1000010,Buffer:=Buffer,Packets:=Packets);
        Capture(PointIndex:=UINT#2,Kind:=USINT#1,Quality:=USINT#2,Value:=LREAL#2.0,NowMs:=ULINT#1000020,NominalDueMs:=ULINT#1000000,SystemUtcMs:=ULINT#1001000,Buffer:=Buffer);
        Policy(Buffer:=Buffer); phaseTicks:=0; Stage:=112;
    END_IF;
112:
    Builder(SliceTestHold:=FALSE,GateOpen:=TRUE,NowMs:=Tick,UnixMs:=ULINT#1002000,GatewayId:='test-gw',BootId:='test-boot',BatchIntervalMs:=UDINT#1,Buffer:=Buffer,Packets:=Packets,Sequence:=Sequence);
    phaseTicks:=phaseTicks+1;
    IF (Buffer.BatchOwners[1].State=2) OR (phaseTicks>500) THEN
        CheckIndex:=48; Check:=(Buffer.BatchOwners[1].Count=1) AND (Buffer.RecordGenerations[firstSlot]<>savedGeneration) AND (FIND(Packets[1].Payload,CONCAT('"value":',TO_STRING(LREAL#2.0,'{0:E16}')))>0) AND (FIND(Packets[1].Payload,CONCAT('"value":',TO_STRING(LREAL#1.0,'{0:E16}')))=0);
        EndBatch(Slot:=UINT#1,Outcome:=USINT#2,Reason:=USINT#0,NowMs:=Tick,Buffer:=Buffer,Packets:=Packets);
        Capture(PointIndex:=UINT#3,Kind:=USINT#1,Quality:=USINT#2,Value:=LREAL#3.0,NowMs:=ULINT#1005010,NominalDueMs:=ULINT#1005000,SystemUtcMs:=ULINT#1006000,Buffer:=Buffer);
        Policy(Buffer:=Buffer); phaseTicks:=0; Stage:=113;
    END_IF;
113:
    Builder(SliceTestHold:=TRUE,GateOpen:=TRUE,NowMs:=Tick,UnixMs:=ULINT#1007000,GatewayId:='test-gw',BootId:='test-boot',BatchIntervalMs:=UDINT#1,Buffer:=Buffer,Packets:=Packets,Sequence:=Sequence);
    phaseTicks:=phaseTicks+1;
    IF Builder.SliceTestPending OR (phaseTicks>500) THEN Stage:=114; END_IF;
114:
    firstSlot:=Buffer.QueueHead[2];
    Builder(SliceTestHold:=FALSE,GateOpen:=FALSE,NowMs:=Tick,UnixMs:=ULINT#1007000,GatewayId:='test-gw',BootId:='test-boot',BatchIntervalMs:=UDINT#1,Buffer:=Buffer,Packets:=Packets,Sequence:=Sequence);
    CheckIndex:=49; Check:=(firstSlot>0) AND (Buffer.QueueHead[2]=firstSlot) AND (Buffer.RecordStates[firstSlot]=1) AND (Buffer.BatchOwners[1].State=0) AND NOT Buffer.CaptureStopped;
    phaseTicks:=0; Stage:=115;
115:
    Builder(GateOpen:=TRUE,NowMs:=Tick,UnixMs:=ULINT#1007000,GatewayId:='test-gw',BootId:='test-boot',BatchIntervalMs:=UDINT#1,Buffer:=Buffer,Packets:=Packets,Sequence:=Sequence);
    phaseTicks:=phaseTicks+1;
    IF (Buffer.BatchOwners[1].State=2) OR (phaseTicks>500) THEN
        CheckIndex:=50; Check:=(Buffer.BatchOwners[1].Count=1) AND (FIND(Packets[1].Payload,CONCAT('"value":',TO_STRING(LREAL#3.0,'{0:E16}')))>0) AND NOT Buffer.CaptureStopped;
        Stage:=116;
    END_IF;
116:
    CheckIndex:=51; Check:=(NG_Quote('')='""') AND (NG_Quote('plain-id')='"plain-id"'); Stage:=117;
117:
    CheckIndex:=52; Check:=NG_Quote('a"b\\c')='"a\\"b\\\\c"'; Stage:=118;
118:
    HashPayload:='a\nb c'; quality:=13;
    firstSlot:=MEMORY_COPY(quality,UDINT#0,HashPayload,UDINT#7,UDINT#1);
    CheckIndex:=53; Check:=(firstSlot=0) AND (NG_Quote(HashPayload)='"a\\nb\\rc"'); Stage:=119;
119:
    CheckIndex:=54; Check:=NG_Quote('a\tb')='"a\\tb"'; Stage:=120;
120:
    EndBatch(Slot:=UINT#1,Outcome:=USINT#2,Reason:=USINT#0,NowMs:=Tick,Buffer:=Buffer,Packets:=Packets);
    Capture(PointIndex:=UINT#1,Kind:=USINT#2,Quality:=USINT#5,Value:=LREAL#0.0,NowMs:=ULINT#1006010,NominalDueMs:=ULINT#0,SystemUtcMs:=ULINT#1006000,Buffer:=Buffer);
    Policy(Buffer:=Buffer); phaseTicks:=0; Stage:=121;
121:
    Builder(GateOpen:=TRUE,NowMs:=Tick,UnixMs:=ULINT#1007000,GatewayId:='test-gw',BootId:='test-boot',BatchIntervalMs:=UDINT#1,Buffer:=Buffer,Packets:=Packets,Sequence:=Sequence);
    phaseTicks:=phaseTicks+1;
    IF (Buffer.BatchOwners[1].State=2) OR (phaseTicks>500) THEN
        CheckIndex:=55; Check:=(FIND(Packets[1].Payload,'"quality":"BAD_TIMEOUT"')>0) AND (FIND(Packets[1].Payload,'"timestamp":1006000')>0) AND (FIND(Packets[1].Payload,'"value":null')>0);
        EndBatch(Slot:=UINT#1,Outcome:=USINT#2,Reason:=USINT#0,NowMs:=Tick,Buffer:=Buffer,Packets:=Packets);
        Capture(PointIndex:=UINT#1,Kind:=USINT#1,Quality:=USINT#2,Value:=LREAL#4.0,NowMs:=ULINT#1010010,NominalDueMs:=ULINT#1010000,SystemUtcMs:=ULINT#1011000,Buffer:=Buffer);
        Policy(Buffer:=Buffer); phaseTicks:=0; Stage:=122;
    END_IF;
122:
    Builder(GateOpen:=TRUE,NowMs:=Tick,UnixMs:=ULINT#1012000,GatewayId:='test-gw',BootId:='test-boot',BatchIntervalMs:=UDINT#1,Buffer:=Buffer,Packets:=Packets,Sequence:=Sequence);
    phaseTicks:=phaseTicks+1;
    IF (Buffer.BatchOwners[1].State=2) OR (phaseTicks>500) THEN
        CheckIndex:=56; Check:=(FIND(Packets[1].Payload,'"quality":"GOOD"')>0) AND (FIND(Packets[1].Payload,'"timestamp":1011000')>0) AND (FIND(Packets[1].Payload,'"value":null')=0);
        Stage:=124;
    END_IF;
124:
    Done:=TRUE;

(* ---- phase1_pipeline_test.st ---- *)
PROGRAM Main
VAR
    Buffer : NG_Buffer;
    EmptyBuffer : NG_Buffer;
    Packets : ARRAY[1..16] OF NG_Packet;
    EmptyPacket : NG_Packet;
    Capture : NG_Capture;
    Source : NG_SourceState;
    SourceResult : NG_SourceResult;
    Policy : NG_ReportPolicy;
    Maintenance : NG_BufferMaintenance;
    Builder : NG_BatchBuilder;
    Delivery : NG_Delivery;
    EndBatch : NG_EndBatch;
    Prune : NG_PruneTerminal;
    StringHash : NG_StringSHA256;
    HashPayload : NG_Json;
    LongPayload : NG_Json;
    LongDigest : STRING[64];
    LongLength : UDINT;
    LongParts : ARRAY[1..64] OF NG_Text;
    Sequence : ULINT;
    Tick : ULINT;
    Stage : INT;
    Scenario : INT := 1;
    Row : INT;
    Rows : INT;
    Passed : UDINT;
    FailedChecks : UDINT;
    Done : BOOL;
    Checks : ARRAY[1..80] OF BOOL;
    CheckIndex : INT;
    Check : BOOL;
    q : ULINT;
    completed : ULINT;
    value : LREAL;
    quality : USINT;
    kind : USINT;
    utc : ULINT;
    pointIndex : UINT;
    i : INT;
    frozen : INT;
    firstSlot : UINT;
    secondSlot : UINT;
    savedId : NG_Id;
    savedPayload : NG_Json;
    savedDigest : STRING[64];
    savedGeneration : UDINT;
    savedSeq : ULINT;
    SubmitAck : BOOL;
    AckId : NG_Id;
    AckStored : BOOL;
    AckRetryable : BOOL;
    Gate : BOOL;
    budget : UDINT;
    BufferBytes : UDINT;
    RecordBytes : UDINT;
    BudgetBytes : UDINT;
    Tx : NG_Bytes;
    Rx : NG_Bytes;
    Values : NG_Json;
    Item : STRING[1024];
    TxPayload : NG_Json;
    DevicesJson : NG_Json;
    Header : STRING[512];
    Samples : ARRAY[1..320] OF NG_Sample;
    Point : NG_Point;
    Sample : NG_Sample;
    phaseTicks : INT;
    AttemptCount : INT;
    StaleCacheValid : BOOL;
    BudgetDigestHeld : BOOL;
    AttemptClasses : ARRAY[1..8] OF USINT;
    SentCount : INT;
    HistoryCount : INT;
    NewCount : INT;
    HashEmptyObject : STRING[64] := '44136fa355b3678a1146ad16f7e8649e94fb4fc21fe77e8310c060f61caaff8a';
END_VAR
IF Done THEN RETURN; END_IF;
Tick:=Tick+20; CheckIndex:=0;
CASE Stage OF
0:
    Buffer:=EmptyBuffer;
    FOR i:=1 TO 16 DO Packets[i]:=EmptyPacket; END_FOR;
    Buffer.ActiveSlot:=1; Buffer.SamplingGeneration:=1; Buffer.LayoutValid:=TRUE;
    Buffer.Configs[1].Generation:=1; Buffer.Configs[1].GatewayId:='test-gw'; Buffer.Configs[1].CaptureBootId:='test-boot';
    Buffer.Configs[1].Config.Version:=1; Buffer.Configs[1].Config.enabled:=TRUE;
    Buffer.Configs[1].Config.maxBatchPoints:=64; Buffer.Configs[1].Config.batchIntervalMs:=1;
    Buffer.Configs[1].Config.DeviceCount:=1; Buffer.Configs[1].Config.PointCount:=64;
    Buffer.Configs[1].Config.Devices[1].deviceId:='device'; Buffer.Configs[1].Config.Devices[1].enabled:=TRUE;
    Buffer.Configs[1].Config.Devices[1].PointStart:=1; Buffer.Configs[1].Config.Devices[1].PointCount:=64;
    FOR i:=1 TO 64 DO
        Buffer.Configs[1].Config.Points[i].pointId:=CONCAT('p',TO_STRING(i,'{0:d}'));
        Buffer.Configs[1].Config.Points[i].enabled:=TRUE; Buffer.Configs[1].Config.Points[i].dataType:='float64';
        Buffer.Configs[1].Config.Points[i].reportMode:='cyclic'; Buffer.Configs[1].Config.Points[i].reportIntervalMs:=5000;
        Buffer.Cursors[i].Enabled:=TRUE; Buffer.Cursors[i].Generation:=1;
    END_FOR;
    IF (Scenario=3) OR (Scenario=4) OR (Scenario=9) THEN Buffer.Configs[1].Config.Points[1].reportMode:='change'; END_IF;
    IF Scenario=3 THEN Buffer.Configs[1].Config.Points[1].deadband:=LREAL#0.5; END_IF;
    IF Scenario=4 THEN Buffer.Configs[1].Config.Points[1].dataType:='bool'; END_IF;
    Row:=0; Rows:=3;
    CASE Scenario OF 2:Rows:=7; 3:Rows:=5; 4,5,6:Rows:=4; 9:Rows:=2; END_CASE;
    IF Scenario<=9 THEN Stage:=1;
    ELSIF Scenario=10 THEN Stage:=10;
    ELSIF Scenario=11 THEN Stage:=30;
    ELSIF Scenario=12 THEN Stage:=50;
    ELSIF Scenario=13 THEN Stage:=60;
    ELSIF Scenario=14 THEN Stage:=70;
    ELSIF Scenario=15 THEN Stage:=80;
    ELSIF Scenario=16 THEN Stage:=90;
    ELSIF Scenario=17 THEN Stage:=100;
    END_IF;
1:
    Row:=Row+1; q:=TO_ULINT(Row-1)*1000; quality:=2; value:=LREAL#10.0; kind:=1;
    CASE Scenario OF
    1:q:=TO_ULINT(Row-1)*5000;
    2:value:=TO_LREAL(Row);
    3:CASE Row OF 1:value:=LREAL#10.0; 2:value:=LREAL#10.5; 3:value:=LREAL#10.6; 4:value:=LREAL#10.9; 5:value:=LREAL#11.2; END_CASE;
    4:IF Row<=2 THEN value:=LREAL#0.0; ELSE value:=LREAL#1.0; END_IF;
    5:IF (Row=2) OR (Row=3) THEN quality:=5; END_IF;
    6:IF Row=1 THEN kind:=2; quality:=1; q:=0; ELSE q:=TO_ULINT(Row-2)*5000; END_IF;
    7:IF Row=3 THEN q:=12000; END_IF;
    END_CASE;
    completed:=q+10;
    IF Scenario=1 THEN
        IF Row=2 THEN completed:=q+8; ELSIF Row=3 THEN completed:=q+11; END_IF;
    ELSIF Scenario=6 THEN
        IF Row=1 THEN completed:=100; ELSIF Row=2 THEN completed:=110; END_IF;
    END_IF;
    IF ((Scenario=8) OR (Scenario=9)) AND (Row=1) THEN Buffer.HighSlot:=28800; Buffer.OwnedCount:=28800; END_IF;
    IF ((Scenario=8) OR (Scenario=9)) AND (Row=2) THEN Buffer.HighSlot:=0; Buffer.OwnedCount:=0; END_IF;
    Capture(PointIndex:=UINT#1,Kind:=kind,Quality:=quality,Value:=value,NowMs:=completed,NominalDueMs:=q,SystemUtcMs:=q+1000,Buffer:=Buffer);
    Policy(Buffer:=Buffer);
    IF Row=Rows THEN Stage:=2; END_IF;
2:
    CheckIndex:=Scenario;
    CASE Scenario OF
    1:Check:=(Buffer.OwnedCount=3) AND (Buffer.Records[1].SampleSeq=1) AND (Buffer.Records[3].SampleSeq=3);
    2:Check:=(Buffer.OwnedCount=2) AND (Buffer.Records[1].SampleSeq=1) AND (Buffer.Records[2].SampleSeq=6);
    3:Check:=(Buffer.OwnedCount=3) AND (Buffer.Records[1].SampleSeq=1) AND (Buffer.Records[2].SampleSeq=3) AND (Buffer.Records[3].SampleSeq=5);
    4:Check:=(Buffer.OwnedCount=2) AND (Buffer.Records[1].Value=LREAL#0.0) AND (Buffer.Records[2].SampleSeq=3);
    5:Check:=(Buffer.OwnedCount=3) AND (Buffer.Records[2].SampleSeq=2) AND (Buffer.Records[3].SampleSeq=4);
    6:Check:=(Buffer.OwnedCount=4) AND (Buffer.ReportCursors[1].NextDue=15000) AND (Buffer.Records[1].Kind=2);
    7:Check:=(Buffer.OwnedCount=2) AND (Buffer.Records[2].SampleSeq=3) AND (Buffer.MissedReportSlotsTotal=1) AND (Buffer.ReportCursors[1].NextDue=15000);
    8:Check:=(Buffer.OwnedCount=1) AND (Buffer.Records[1].SampleSeq=2) AND (Buffer.KnownUnsentEventsTotal=1) AND (Buffer.EnqueueRejectedAttemptsTotal=1) AND (Buffer.ReportCursors[1].NextDue=5000) AND (Buffer.MissedReportSlotsTotal=0);
    9:Check:=(Buffer.OwnedCount=1) AND (Buffer.Records[1].SampleSeq=2) AND (Buffer.KnownUnsentEventsTotal=1);
    END_CASE;
    Scenario:=Scenario+1; Stage:=0;
10:
    (* Same point's two physical events remain distinct across builder windows. *)
    Capture(PointIndex:=UINT#1,Kind:=USINT#1,Quality:=USINT#2,Value:=LREAL#10.0,NowMs:=ULINT#10,NominalDueMs:=ULINT#0,SystemUtcMs:=ULINT#1000,Buffer:=Buffer);
    Policy(Buffer:=Buffer);
    Capture(PointIndex:=UINT#1,Kind:=USINT#1,Quality:=USINT#2,Value:=LREAL#20.0,NowMs:=ULINT#5010,NominalDueMs:=ULINT#5000,SystemUtcMs:=ULINT#6000,Buffer:=Buffer);
    Policy(Buffer:=Buffer); Stage:=11; phaseTicks:=0;
11:
    Builder(GateOpen:=TRUE,NowMs:=Tick,UnixMs:=ULINT#10000,GatewayId:='test-gw',BootId:='test-boot',BatchIntervalMs:=UDINT#1,Buffer:=Buffer,Packets:=Packets,Sequence:=Sequence);
    frozen:=0; FOR i:=1 TO 16 DO IF Buffer.BatchOwners[i].State=2 THEN frozen:=frozen+1; END_IF; END_FOR;
    phaseTicks:=phaseTicks+1;
    IF (frozen=2) OR (phaseTicks>200) THEN
        CheckIndex:=10; Check:=(frozen=2) AND (Buffer.BatchOwners[1].Count=1) AND (Buffer.BatchOwners[2].Count=1) AND (Packets[1].MessageId<>Packets[2].MessageId) AND (Buffer.Records[Buffer.BatchRefs[1]].SampleSeq=1) AND (Buffer.Records[Buffer.BatchRefs[65]].SampleSeq=2);
        savedId:=Packets[1].MessageId; savedPayload:=Packets[1].Payload; savedDigest:=Buffer.BatchOwners[1].Digest;
        savedGeneration:=Buffer.BatchGenerations[1];
        Packets[1].WasSent:=TRUE; Packets[2].WasSent:=TRUE;
        AckId:=Packets[2].MessageId; AckStored:=TRUE; AckRetryable:=FALSE; SubmitAck:=TRUE; Stage:=12; phaseTicks:=0;
    END_IF;
12:
    Delivery(GateOpen:=FALSE,NowMs:=Tick,GatewayId:='test-gw',BootId:='test-boot',SubmitAck:=SubmitAck,AckMessageId:=AckId,AckStored:=AckStored,AckRetryable:=AckRetryable,AckCodes:='',Buffer:=Buffer,Packets:=Packets);
    SubmitAck:=FALSE;
    phaseTicks:=phaseTicks+1;
    IF NOT Delivery.AckBusy OR (phaseTicks>200) THEN
        CheckIndex:=11; Check:=(Buffer.StoredConfirmedEventsTotal=1) AND (Buffer.OwnedCount=1) AND (Packets[1].Payload=savedPayload) AND (Buffer.ReportCursors[1].LastSeq=2);
        AckId:=savedId; SubmitAck:=TRUE; Stage:=13; phaseTicks:=0;
    END_IF;
13:
    Delivery(GateOpen:=FALSE,NowMs:=Tick,GatewayId:='test-gw',BootId:='test-boot',SubmitAck:=SubmitAck,AckMessageId:=AckId,AckStored:=TRUE,AckRetryable:=FALSE,AckCodes:='',Buffer:=Buffer,Packets:=Packets);
    SubmitAck:=FALSE;
    phaseTicks:=phaseTicks+1;
    IF NOT Delivery.AckBusy OR (phaseTicks>200) THEN
        CheckIndex:=12; Check:=(Buffer.StoredConfirmedEventsTotal=2) AND (Buffer.OwnedCount=0) AND (Buffer.ReportCursors[1].LastSeq=2);
        Capture(PointIndex:=UINT#1,Kind:=USINT#1,Quality:=USINT#2,Value:=LREAL#20.0,NowMs:=ULINT#6010,NominalDueMs:=ULINT#6000,SystemUtcMs:=ULINT#7000,Buffer:=Buffer); Policy(Buffer:=Buffer);
        Stage:=14;
    END_IF;
14:
    CheckIndex:=13; Check:=(Buffer.OwnedCount=0) AND (Buffer.PolicyFilteredEventsTotal=1) AND (Buffer.ReportCursors[1].LastSeq=2);
    Capture(PointIndex:=UINT#1,Kind:=USINT#1,Quality:=USINT#2,Value:=LREAL#20.0,NowMs:=ULINT#10010,NominalDueMs:=ULINT#10000,SystemUtcMs:=ULINT#11000,Buffer:=Buffer); Policy(Buffer:=Buffer);
    Stage:=15; phaseTicks:=0;
15:
    Builder(GateOpen:=TRUE,NowMs:=Tick,UnixMs:=ULINT#12000,GatewayId:='test-gw',BootId:='test-boot',BatchIntervalMs:=UDINT#1,Buffer:=Buffer,Packets:=Packets,Sequence:=Sequence);
    phaseTicks:=phaseTicks+1;
    IF (Buffer.BatchOwners[1].State=2) OR (phaseTicks>200) THEN
        CheckIndex:=14; Check:=(Buffer.BatchGenerations[1]>savedGeneration) AND (Packets[1].MessageId<>savedId);
        AckId:=savedId; SubmitAck:=TRUE; Stage:=16;
    END_IF;
16:
    Delivery(GateOpen:=FALSE,NowMs:=Tick,GatewayId:='test-gw',BootId:='test-boot',SubmitAck:=SubmitAck,AckMessageId:=AckId,AckStored:=TRUE,AckRetryable:=FALSE,AckCodes:='',Buffer:=Buffer,Packets:=Packets);
    SubmitAck:=FALSE;
    CheckIndex:=15; Check:=(Buffer.OwnedCount=1) AND (Buffer.BatchOwners[1].State=2) AND (Buffer.StoredConfirmedEventsTotal=2);
    Packets[1].WasSent:=TRUE; savedId:=Packets[1].MessageId; savedPayload:=Packets[1].Payload;
    EndBatch(Slot:=UINT#1,Outcome:=USINT#4,Reason:=USINT#5,NowMs:=Tick,Buffer:=Buffer,Packets:=Packets);
    AckId:=savedId; SubmitAck:=TRUE; Stage:=17;
17:
    Delivery(GateOpen:=FALSE,NowMs:=Tick,GatewayId:='test-gw',BootId:='test-boot',SubmitAck:=SubmitAck,AckMessageId:=AckId,AckStored:=TRUE,AckRetryable:=FALSE,AckCodes:='',Buffer:=Buffer,Packets:=Packets);
    SubmitAck:=FALSE;
    CheckIndex:=16; Check:=(Buffer.UncertainDeliveryEventsTotal=1) AND (Buffer.LateStoredEventsTotal=1) AND (Buffer.StoredConfirmedEventsTotal=3) AND (Buffer.OwnedCount=0);
    SubmitAck:=TRUE; Stage:=18;
18:
    Delivery(GateOpen:=FALSE,NowMs:=Tick,GatewayId:='test-gw',BootId:='test-boot',SubmitAck:=SubmitAck,AckMessageId:=AckId,AckStored:=TRUE,AckRetryable:=FALSE,AckCodes:='',Buffer:=Buffer,Packets:=Packets);
    SubmitAck:=FALSE;
    CheckIndex:=17; Check:=(Buffer.LateStoredEventsTotal=1) AND (Buffer.StoredConfirmedEventsTotal=3);
    Stage:=20;
20:
    (* Time invalid rejects only this selected event; prior admitted owner stays. *)
    Capture(PointIndex:=UINT#1,Kind:=USINT#1,Quality:=USINT#2,Value:=LREAL#30.0,NowMs:=ULINT#15010,NominalDueMs:=ULINT#15000,SystemUtcMs:=ULINT#16000,Buffer:=Buffer); Policy(Buffer:=Buffer);
    savedSeq:=Buffer.Records[Buffer.QueueHead[2]].SampleSeq;
    Capture(PointIndex:=UINT#1,Kind:=USINT#1,Quality:=USINT#2,Value:=LREAL#40.0,NowMs:=ULINT#20010,NominalDueMs:=ULINT#20000,SystemUtcMs:=ULINT#0,Buffer:=Buffer); Policy(Buffer:=Buffer);
    CheckIndex:=18; Check:=(Buffer.OwnedCount=1) AND (Buffer.TimeInvalidEventsTotal=1) AND (Buffer.KnownUnsentEventsTotal=1) AND (Buffer.Records[Buffer.QueueHead[2]].SampleSeq=savedSeq);
    Capture(PointIndex:=UINT#1,Kind:=USINT#1,Quality:=USINT#2,Value:=LREAL#40.0,NowMs:=ULINT#21010,NominalDueMs:=ULINT#21000,SystemUtcMs:=ULINT#22000,Buffer:=Buffer); Policy(Buffer:=Buffer);
    Stage:=21;
21:
    CheckIndex:=19; Check:=(Buffer.OwnedCount=2) AND (Buffer.ReportCursors[1].LastSeq=7);
    Buffer.ActiveSlot:=2; Buffer.Configs[2].Generation:=2; Buffer.SamplingGeneration:=2;
    Maintenance(GateOpen:=FALSE,NowMs:=Tick,Buffer:=Buffer,Packets:=Packets);
    Stage:=22;
22:
    CheckIndex:=20; Check:=(Buffer.OwnedCount=2) AND (Buffer.Configs[1].References=2) AND (Buffer.Records[Buffer.QueueHead[2]].ConfigSlot=1);
    Buffer.ActiveSlot:=1; Buffer.SamplingGeneration:=1;
    Maintenance(GateOpen:=TRUE,NowMs:=Tick,Buffer:=Buffer,Packets:=Packets);
    Capture(PointIndex:=UINT#2,Kind:=USINT#1,Quality:=USINT#2,Value:=LREAL#1.0,NowMs:=ULINT#10,NominalDueMs:=ULINT#0,SystemUtcMs:=ULINT#1000,Buffer:=Buffer); Policy(Buffer:=Buffer);
    Stage:=23;
23:
    CheckIndex:=21; Check:=(Buffer.QueueHead[1]<>0) AND (Buffer.QueueHead[2]<>0) AND (Buffer.Records[Buffer.QueueHead[2]].SampleSeq>Buffer.Watermark);
    HashPayload:='abc'; Stage:=24;
24:
    StringHash(Execute:=TRUE,Length:=UDINT#3,Payload:=HashPayload);
    IF StringHash.Done THEN
        CheckIndex:=22; Check:=StringHash.Digest='ba7816bf8f01cfea414140de5dae2223b00361a396177a9cb410ff61f20015ad'; Stage:=25;
    END_IF;
25:
    RecordBytes:=SIZEOF(Buffer.Scratch); BufferBytes:=SIZEOF(Buffer);
    budget:=SIZEOF(Packets)+SIZEOF(Samples)+SIZEOF(Values)+SIZEOF(Item)+SIZEOF(TxPayload)+SIZEOF(EmptyPacket)+SIZEOF(Sample)+SIZEOF(Point)+SIZEOF(Tx)+SIZEOF(Rx)+SIZEOF(DevicesJson)+SIZEOF(Header)+UDINT#16384+UDINT#135680+UDINT#65536;
    BudgetBytes:=BufferBytes+budget;
    CheckIndex:=23; Check:=(RecordBytes=72) AND (BudgetBytes<=4194304); Stage:=26;
26:
    Scenario:=11; Stage:=0;
30:
    FOR i:=1 TO 16 DO
        Capture(PointIndex:=TO_UINT(i),Kind:=USINT#1,Quality:=USINT#2,Value:=LREAL#-1.2345678901234567E300,NowMs:=ULINT#10,NominalDueMs:=ULINT#0,SystemUtcMs:=ULINT#9007199254740991,Buffer:=Buffer);
    END_FOR;
    Policy(Buffer:=Buffer); Buffer.QueueHead[2]:=0; Buffer.QueueTail[2]:=0;
    FOR i:=1 TO 16 DO
        Packets[i].Payload:='{}'; Packets[i].Length:=2; Packets[i].MessageId:=CONCAT('fixture-',TO_STRING(i,'{0:d}'));
        Buffer.BatchGenerations[i]:=1; Buffer.BatchOwners[i].State:=2; Buffer.BatchOwners[i].Count:=1;
        Buffer.BatchOwners[i].OrderSeq:=TO_ULINT(i); Buffer.BatchOwners[i].ConfigSlot:=1;
        Buffer.BatchOwners[i].Digest:=HashEmptyObject; Buffer.BatchOwners[i].Category:=1;
        IF i>8 THEN Buffer.BatchOwners[i].Category:=2; END_IF;
        Buffer.BatchRefs[(i-1)*64+1]:=TO_UINT(i); Buffer.BatchRefGenerations[(i-1)*64+1]:=Buffer.RecordGenerations[i];
        Buffer.RecordStates[i]:=2;
    END_FOR;
    AttemptCount:=0; phaseTicks:=0; Stage:=31;
31:
    Delivery(GateOpen:=TRUE,NowMs:=Tick,GatewayId:='test-gw',BootId:='test-boot',SubmitAck:=FALSE,AckMessageId:='',AckStored:=FALSE,AckRetryable:=FALSE,AckCodes:='',Buffer:=Buffer,Packets:=Packets);
    phaseTicks:=phaseTicks+1;
    IF Delivery.SendSlot>0 THEN
        firstSlot:=Delivery.SendSlot; AttemptCount:=AttemptCount+1; AttemptClasses[AttemptCount]:=Buffer.BatchOwners[firstSlot].Category;
        Packets[firstSlot].WasSent:=TRUE; Packets[firstSlot].Attempts:=1; Packets[firstSlot].RetryAtMs:=Tick+30000;
        Buffer.NextSendAt:=Tick+334; Buffer.PreferSend:=USINT#3-Buffer.BatchOwners[firstSlot].Category;
    END_IF;
    IF (AttemptCount=8) OR (phaseTicks>500) THEN
        SentCount:=0; HistoryCount:=0; NewCount:=0;
        FOR i:=1 TO 16 DO
            IF Packets[i].WasSent THEN SentCount:=SentCount+1;
                IF Buffer.BatchOwners[i].Category=1 THEN HistoryCount:=HistoryCount+1; ELSE NewCount:=NewCount+1; END_IF;
            END_IF;
        END_FOR;
        CheckIndex:=24; Check:=(AttemptCount=8) AND (SentCount=8) AND (HistoryCount=4) AND (NewCount=4);
        FOR i:=2 TO 8 DO Check:=Check AND (AttemptClasses[i]<>AttemptClasses[i-1]); END_FOR;
        Stage:=32; phaseTicks:=0;
    END_IF;
32:
    Delivery(GateOpen:=TRUE,NowMs:=Tick,GatewayId:='test-gw',BootId:='test-boot',SubmitAck:=FALSE,AckMessageId:='',AckStored:=FALSE,AckRetryable:=FALSE,AckCodes:='',Buffer:=Buffer,Packets:=Packets);
    phaseTicks:=phaseTicks+1;
    IF phaseTicks=30 THEN CheckIndex:=25; Check:=(Delivery.SendSlot=0) AND (Buffer.OwnedCount=16); Tick:=Tick+31000; Stage:=33; phaseTicks:=0; END_IF;
33:
    Delivery(GateOpen:=TRUE,NowMs:=Tick,GatewayId:='test-gw',BootId:='test-boot',SubmitAck:=FALSE,AckMessageId:='',AckStored:=FALSE,AckRetryable:=FALSE,AckCodes:='',Buffer:=Buffer,Packets:=Packets);
    phaseTicks:=phaseTicks+1;
    IF (Delivery.SendSlot>0) OR (phaseTicks>100) THEN
        CheckIndex:=26; Check:=FALSE;
        IF Delivery.SendSlot>0 THEN Check:=Packets[Delivery.SendSlot].WasSent; END_IF;
        firstSlot:=Delivery.SendSlot; AckId:=Packets[firstSlot].MessageId; SubmitAck:=TRUE; phaseTicks:=0; Stage:=34;
    END_IF;
34:
    Delivery(GateOpen:=FALSE,NowMs:=Tick,GatewayId:='test-gw',BootId:='test-boot',SubmitAck:=SubmitAck,AckMessageId:=AckId,AckStored:=FALSE,AckRetryable:=TRUE,AckCodes:='STORAGE_ERROR',Buffer:=Buffer,Packets:=Packets);
    SubmitAck:=FALSE; phaseTicks:=phaseTicks+1;
    IF NOT Delivery.AckBusy OR (phaseTicks>100) THEN
        CheckIndex:=27; Check:=(Packets[firstSlot].RetryAtMs>=Tick+60000) AND (Buffer.StoredConfirmedEventsTotal=0) AND (Buffer.IsolatedEventsTotal=0);
        savedSeq:=Packets[firstSlot].RetryAtMs; Maintenance(GateOpen:=FALSE,NowMs:=Tick,Buffer:=Buffer,Packets:=Packets);
        Maintenance(GateOpen:=TRUE,NowMs:=Tick,Buffer:=Buffer,Packets:=Packets);
        Stage:=35;
    END_IF;
35:
    CheckIndex:=28; Check:=(Packets[firstSlot].RetryAtMs=savedSeq) AND (Packets[firstSlot].Attempts=1);
    AckId:=Packets[2].MessageId; Packets[2].WasSent:=TRUE; SubmitAck:=TRUE; Stage:=36; phaseTicks:=0;
36:
    Delivery(GateOpen:=FALSE,NowMs:=Tick,GatewayId:='test-gw',BootId:='test-boot',SubmitAck:=SubmitAck,AckMessageId:=AckId,AckStored:=FALSE,AckRetryable:=FALSE,AckCodes:='VALIDATION_ERROR',Buffer:=Buffer,Packets:=Packets);
    SubmitAck:=FALSE; phaseTicks:=phaseTicks+1;
    IF NOT Delivery.AckBusy OR (phaseTicks>100) THEN
        CheckIndex:=29; Check:=(Buffer.BatchOwners[2].State=3) AND (Buffer.IsolatedEventsTotal=1) AND Packets[2].Dead;
        SubmitAck:=TRUE; Stage:=37; phaseTicks:=0;
    END_IF;
37:
    Delivery(GateOpen:=FALSE,NowMs:=Tick,GatewayId:='test-gw',BootId:='test-boot',SubmitAck:=SubmitAck,AckMessageId:=AckId,AckStored:=TRUE,AckRetryable:=FALSE,AckCodes:='',Buffer:=Buffer,Packets:=Packets);
    SubmitAck:=FALSE; phaseTicks:=phaseTicks+1;
    IF NOT Delivery.AckBusy OR (phaseTicks>100) THEN
        CheckIndex:=30; Check:=(Buffer.IsolatedEventsTotal=1) AND (Buffer.StoredConfirmedEventsTotal=0) AND (Buffer.ConflictingAcksTotal=1);
        FOR i:=1 TO 6 DO EndBatch(Slot:=TO_UINT(i),Outcome:=USINT#3,Reason:=USINT#8,NowMs:=Tick,Buffer:=Buffer,Packets:=Packets); END_FOR;
        Stage:=38;
    END_IF;
38:
    Maintenance(GateOpen:=FALSE,NowMs:=Tick,Buffer:=Buffer,Packets:=Packets);
    Maintenance(GateOpen:=FALSE,NowMs:=Tick,Buffer:=Buffer,Packets:=Packets);
    frozen:=0; FOR i:=1 TO 16 DO IF Buffer.BatchOwners[i].State=3 THEN frozen:=frozen+1; END_IF; END_FOR;
    CheckIndex:=31; Check:=(frozen=4) AND (Buffer.IsolatedEventsTotal=6) AND (Buffer.DeadPrunedBatchesTotal=2) AND (Buffer.OwnedCount=16);
    Prune(Index:=UINT#1,Buffer:=Buffer); Stage:=39;
39:
    CheckIndex:=32; Check:=(Buffer.IsolatedEventsTotal=6) AND (Buffer.TombstonePrunedBatchesTotal=1) AND (Buffer.OwnedCount=15) AND Buffer.DetailTruncated;
    Packets[15].WasSent:=TRUE; Packets[15].Payload:='{"changed":true}'; Packets[15].Length:=16;
    AckId:=Packets[15].MessageId; SubmitAck:=TRUE; Stage:=40; phaseTicks:=0;
40:
    Delivery(GateOpen:=FALSE,NowMs:=Tick,GatewayId:='test-gw',BootId:='test-boot',SubmitAck:=SubmitAck,AckMessageId:=AckId,AckStored:=TRUE,AckRetryable:=FALSE,AckCodes:='',Buffer:=Buffer,Packets:=Packets);
    SubmitAck:=FALSE; phaseTicks:=phaseTicks+1;
    IF NOT Delivery.AckBusy OR (phaseTicks>100) THEN
        CheckIndex:=33; Check:=Buffer.CaptureStopped AND NOT Buffer.AccountingComplete AND (Buffer.CorruptBatchesTotal=1) AND (Buffer.StoredConfirmedEventsTotal=0) AND (Buffer.UncertainDeliveryEventsTotal=1);
        Scenario:=12; Stage:=0;
    END_IF;
50:
    FOR i:=1 TO 8 DO Capture(PointIndex:=TO_UINT(i),Kind:=USINT#1,Quality:=USINT#2,Value:=TO_LREAL(i),NowMs:=ULINT#10,NominalDueMs:=ULINT#0,SystemUtcMs:=ULINT#1000,Buffer:=Buffer); END_FOR;
    Policy(Buffer:=Buffer);
    Builder(GateOpen:=TRUE,NowMs:=Tick,UnixMs:=ULINT#2000,GatewayId:='test-gw',BootId:='test-boot',BatchIntervalMs:=UDINT#1,Buffer:=Buffer,Packets:=Packets,Sequence:=Sequence);
    Stage:=51;
51:
    Builder(GateOpen:=FALSE,NowMs:=Tick,UnixMs:=ULINT#0,GatewayId:='test-gw',BootId:='test-boot',BatchIntervalMs:=UDINT#1,Buffer:=Buffer,Packets:=Packets,Sequence:=Sequence);
    CheckIndex:=34; Check:=(Buffer.OwnedCount=8) AND (Buffer.BatchOwners[1].State=0) AND (Buffer.Records[Buffer.QueueHead[2]].SampleSeq=1) AND (Buffer.Records[Buffer.QueueTail[2]].SampleSeq=8) AND (Buffer.KnownUnsentEventsTotal=0);
    Scenario:=13; Stage:=0;
60:
    (* Mutating a frozen dictionary requires a new generation, as in the real allocator. *)
    Buffer.Configs[1].Generation:=2;
    Buffer.Configs[1].Config.DeviceCount:=2; Buffer.Configs[1].Config.Devices[1].PointCount:=32;
    Buffer.Configs[1].Config.Devices[1].deviceId:='dddddddddddddddddddddddddddddddddddddddddddddddddddddddddddddddd';
    Buffer.Configs[1].Config.Devices[2].deviceId:='eeeeeeeeeeeeeeeeeeeeeeeeeeeeeeeeeeeeeeeeeeeeeeeeeeeeeeeeeeeeeeee';
    Buffer.Configs[1].Config.Devices[2].enabled:=TRUE; Buffer.Configs[1].Config.Devices[2].PointStart:=33; Buffer.Configs[1].Config.Devices[2].PointCount:=32;
    FOR i:=1 TO 64 DO
        Buffer.Configs[1].Config.Points[i].pointId:=CONCAT('pppppppppppppppppppppppppppppppppppppppppppppppppppppppppppppp',TO_STRING(i,'{0:d}'));
        Capture(PointIndex:=TO_UINT(i),Kind:=USINT#1,Quality:=USINT#2,Value:=LREAL#-1.2345678901234567E300,NowMs:=ULINT#10,NominalDueMs:=ULINT#0,SystemUtcMs:=ULINT#9007199254740991,Buffer:=Buffer);
    END_FOR;
    Policy(Buffer:=Buffer); Stage:=61; phaseTicks:=0;
61:
    Builder(GateOpen:=TRUE,NowMs:=Tick,UnixMs:=ULINT#2000,GatewayId:='test-gw',BootId:='test-boot',BatchIntervalMs:=UDINT#1,Buffer:=Buffer,Packets:=Packets,Sequence:=Sequence);
    phaseTicks:=phaseTicks+1; frozen:=0; SentCount:=0;
    FOR i:=1 TO 16 DO IF Buffer.BatchOwners[i].State=2 THEN frozen:=frozen+1; SentCount:=SentCount+TO_INT(Buffer.BatchOwners[i].Count); END_IF; END_FOR;
    IF (SentCount=64) OR (phaseTicks>500) THEN
        CheckIndex:=35; Check:=(SentCount=64) AND (frozen>=1) AND (Buffer.OwnedCount=64) AND (Buffer.QueueHead[2]=0);
        FOR i:=1 TO 16 DO IF Buffer.BatchOwners[i].State=2 THEN Check:=Check AND (Packets[i].Length<=16380) AND (Packets[i].Length=TO_UDINT(LEN(Packets[i].Payload))) AND (RIGHT(Packets[i].Payload,2)=']}') AND (Buffer.BatchOwners[i].Count<=64); END_IF; END_FOR;
        LongPayload:=Packets[1].Payload; LongDigest:=Buffer.BatchOwners[1].Digest; LongLength:=Packets[1].Length;
        FOR i:=1 TO 64 DO
            LongParts[i]:='';
            IF (i-1)*256<LEN(LongPayload) THEN LongParts[i]:=MID(LongPayload,MIN(256,LEN(LongPayload)-(i-1)*256),(i-1)*256+1); END_IF;
        END_FOR;
        Stage:=62;
    END_IF;
62:
    Maintenance(GateOpen:=FALSE,NowMs:=ULINT#900010,Buffer:=Buffer,Packets:=Packets);
    Maintenance(GateOpen:=FALSE,NowMs:=ULINT#900010,Buffer:=Buffer,Packets:=Packets);
    CheckIndex:=36; Check:=(Buffer.KnownUnsentEventsTotal=64) AND (Buffer.OwnedCount=0) AND (Buffer.UncertainDeliveryEventsTotal=0);
    Scenario:=14; Stage:=0;
70:
    FOR i:=1 TO 64 DO Capture(PointIndex:=TO_UINT(i),Kind:=USINT#1,Quality:=USINT#2,Value:=TO_LREAL(i),NowMs:=ULINT#10,NominalDueMs:=ULINT#0,SystemUtcMs:=ULINT#1000,Buffer:=Buffer); END_FOR;
    Policy(Buffer:=Buffer); Maintenance(GateOpen:=FALSE,NowMs:=ULINT#900010,Buffer:=Buffer,Packets:=Packets);
    CheckIndex:=37; Check:=(Buffer.KnownUnsentEventsTotal=64) AND (Buffer.OwnedCount=0) AND (Buffer.Configs[1].References=0) AND (Buffer.GapRecordsTotal=64);
    Scenario:=15; Stage:=0; Row:=0;
80:
    FOR i:=1 TO 64 DO
        q:=Buffer.NextSampleSeq*5000;
        Capture(PointIndex:=UINT#1,Kind:=USINT#1,Quality:=USINT#2,Value:=TO_LREAL(Buffer.NextSampleSeq),NowMs:=q+10,NominalDueMs:=q,SystemUtcMs:=q+1000,Buffer:=Buffer);
    END_FOR;
    Policy(Buffer:=Buffer);
    IF Buffer.OwnedCount=28800 THEN Stage:=81; END_IF;
81:
    savedSeq:=Buffer.Records[Buffer.QueueHead[2]].SampleSeq;
    FOR i:=1 TO 64 DO
        q:=Buffer.NextSampleSeq*5000;
        Capture(PointIndex:=UINT#1,Kind:=USINT#1,Quality:=USINT#2,Value:=TO_LREAL(Buffer.NextSampleSeq),NowMs:=q+10,NominalDueMs:=q,SystemUtcMs:=q+1000,Buffer:=Buffer);
    END_FOR;
    Maintenance(GateOpen:=FALSE,NowMs:=ULINT#0,Buffer:=Buffer,Packets:=Packets); Policy(Buffer:=Buffer);
    CheckIndex:=38; Check:=(Buffer.OwnedCount=28800) AND (Buffer.KnownUnsentEventsTotal=64) AND (Buffer.EnqueueRejectedAttemptsTotal=0) AND (Buffer.Records[Buffer.QueueHead[2]].SampleSeq=savedSeq+64) AND (Buffer.Configs[1].References=28800);
    Stage:=82;
82:
    firstSlot:=Buffer.QueueHead[2]; Buffer.QueueHead[2]:=Buffer.FreeSlots[firstSlot];
    Packets[1].MessageId:='pressure-sent'; Packets[1].Payload:='{}'; Packets[1].Length:=2; Packets[1].WasSent:=TRUE;
    Buffer.BatchOwners[1].State:=2; Buffer.BatchOwners[1].Count:=1; Buffer.BatchOwners[1].Category:=2;
    Buffer.BatchOwners[1].ConfigSlot:=1; Buffer.BatchOwners[1].OrderSeq:=Buffer.Records[firstSlot].SampleSeq;
    Buffer.BatchOwners[1].Digest:=HashEmptyObject; Buffer.BatchRefs[1]:=firstSlot;
    Buffer.BatchRefGenerations[1]:=Buffer.RecordGenerations[firstSlot]; Buffer.RecordStates[firstSlot]:=2;
    q:=Buffer.NextSampleSeq*5000;
    Capture(PointIndex:=UINT#1,Kind:=USINT#1,Quality:=USINT#2,Value:=LREAL#1.0,NowMs:=q+10,NominalDueMs:=q,SystemUtcMs:=q+1000,Buffer:=Buffer);
    Maintenance(GateOpen:=FALSE,NowMs:=ULINT#0,Buffer:=Buffer,Packets:=Packets); Policy(DeferCapacity:=TRUE,Buffer:=Buffer); Stage:=83;
83:
    CheckIndex:=41; Check:=(Buffer.OwnedCount=28800) AND (Buffer.UncertainDeliveryEventsTotal=1) AND (Buffer.TombstonePrunedBatchesTotal=1) AND (Buffer.KnownUnsentEventsTotal=64) AND (Buffer.IngressCount=0) AND (Buffer.Configs[1].References=28800);
    Scenario:=16; Stage:=0;
90:
    Buffer.Configs[1].Config.Points[1].staleAfterMs:=3000;
    Buffer.Cursors[1].Enabled:=FALSE;
    Source(Index:=UINT#1,Enabled:=TRUE,NowMs:=ULINT#1000,UnixMs:=ULINT#2000,StaleAfterMs:=UDINT#3000,CheckStale:=TRUE,Samples:=Samples,Buffer:=Buffer);
    StaleCacheValid:=Buffer.SourceStaleDue[1]=4000;
    FOR i:=0 TO 2 DO
        q:=ULINT#1010+TO_ULINT(i)*1000;
        SourceResult(Index:=UINT#1,Value:=LREAL#0.0,Quality:='BAD_TIMEOUT',NowMs:=q,UnixMs:=q+1000,NominalDueMs:=q-10,ConfigSlot:=UINT#1,ConfigGeneration:=UDINT#1,SamplingGeneration:=ULINT#1,Samples:=Samples,Buffer:=Buffer);
        StaleCacheValid:=StaleCacheValid AND (Buffer.SourceStaleDue[1]=q+3000);
        Source(Index:=UINT#1,Enabled:=TRUE,NowMs:=q,UnixMs:=q+1000,StaleAfterMs:=UDINT#3000,CheckStale:=TRUE,Samples:=Samples,Buffer:=Buffer);
    END_FOR;
    Source(Index:=UINT#1,Enabled:=TRUE,NowMs:=ULINT#6009,UnixMs:=ULINT#7009,StaleAfterMs:=UDINT#3000,CheckStale:=TRUE,Samples:=Samples,Buffer:=Buffer);
    StaleCacheValid:=StaleCacheValid AND (Buffer.SourceStaleDue[1]=6010);
    savedSeq:=Buffer.CapturedEventsTotal;
    FOR i:=1 TO 100 DO Source(Index:=UINT#1,Enabled:=TRUE,NowMs:=ULINT#6010+TO_ULINT(i-1),UnixMs:=ULINT#7010+TO_ULINT(i-1),StaleAfterMs:=UDINT#3000,CheckStale:=TRUE,Samples:=Samples,Buffer:=Buffer); END_FOR;
    Policy(Buffer:=Buffer); Stage:=91;
91:
    CheckIndex:=39; Check:=StaleCacheValid AND (Buffer.SourceStaleDue[1]=0) AND (savedSeq=4) AND (Buffer.CapturedEventsTotal=5) AND (Buffer.OwnedCount=3) AND (Buffer.PolicyFilteredEventsTotal=2) AND (Samples[1].Quality='STALE') AND (Samples[1].LastGoodMs=0);
    Capture(PointIndex:=UINT#1,Kind:=USINT#1,Quality:=USINT#2,Value:=LREAL#1.0,NowMs:=ULINT#10010,NominalDueMs:=ULINT#10000,SystemUtcMs:=ULINT#11000,Buffer:=Buffer);
    Buffer.ActiveSlot:=2; Buffer.SamplingGeneration:=2; Policy(Buffer:=Buffer); Stage:=92;
92:
    CheckIndex:=40; Check:=(Buffer.UndecidedLostEventsTotal=1) AND (Buffer.EligibleEventsTotal=3) AND (Buffer.PolicyFilteredEventsTotal=2) AND (Buffer.OwnedCount=3) AND NOT Buffer.AccountingComplete AND (Buffer.Gaps[Buffer.GapIndex].Reason=2);
    Stage:=93;
93:
    HashPayload:=LongPayload;
    StringHash(Execute:=FALSE,Length:=LongLength,DeadlineUs:=ULINT#1,Payload:=HashPayload);
    StringHash(Execute:=TRUE,Length:=LongLength,DeadlineUs:=ULINT#1,Payload:=HashPayload);
    BudgetDigestHeld:=StringHash.Busy AND NOT StringHash.Done;
    phaseTicks:=0; Stage:=94;
94:
    (* An expired absolute deadline may not advance an in-progress digest.
       Fresh bounded slices must still produce the independent long vector. *)
    savedDigest:=StringHash.Digest;
    StringHash(Execute:=TRUE,Length:=LongLength,DeadlineUs:=ULINT#1,Payload:=HashPayload);
    BudgetDigestHeld:=BudgetDigestHeld AND (savedDigest=StringHash.Digest) AND StringHash.Busy AND NOT StringHash.Done;
    StringHash(Execute:=TRUE,Length:=LongLength,DeadlineUs:=GET_MICROSECONDS(TRUE)+ULINT#250,Payload:=HashPayload);
    phaseTicks:=phaseTicks+1;
    IF StringHash.Done OR (phaseTicks>2000) THEN Stage:=95; END_IF;
95:
    CheckIndex:=42; Check:=StringHash.Done AND NOT StringHash.Error AND (StringHash.Digest=LongDigest);
    Stage:=96;
96:
    CheckIndex:=43; Check:=BudgetDigestHeld;
    Stage:=97;
97:
    Scenario:=17; Stage:=0;
100:
    Buffer.Configs[1].Config.Devices[1].deviceId:='new"device';
    Capture(PointIndex:=UINT#1,Kind:=USINT#1,Quality:=USINT#2,Value:=LREAL#1.0,NowMs:=ULINT#10,NominalDueMs:=ULINT#0,SystemUtcMs:=ULINT#1000,Buffer:=Buffer);
    Policy(Buffer:=Buffer); phaseTicks:=0; Stage:=101;
101:
    Builder(GateOpen:=TRUE,NowMs:=Tick,UnixMs:=ULINT#2000,GatewayId:='test-gw',BootId:='test-boot',BatchIntervalMs:=UDINT#1,Buffer:=Buffer,Packets:=Packets,Sequence:=Sequence);
    phaseTicks:=phaseTicks+1;
    IF (Buffer.BatchOwners[1].State=2) OR (phaseTicks>500) THEN
        CheckIndex:=44; Check:=(Buffer.BatchOwners[1].Count=1) AND (FIND(Packets[1].Payload,CONCAT('"deviceId":',NG_Quote('new"device')))>0);
        EndBatch(Slot:=UINT#1,Outcome:=USINT#2,Reason:=USINT#0,NowMs:=Tick,Buffer:=Buffer,Packets:=Packets);
        Stage:=102;
    END_IF;
102:
    Buffer.Configs[1].Generation:=2; Buffer.Configs[1].Config.Devices[1].deviceId:='changed"device';
    Capture(PointIndex:=UINT#1,Kind:=USINT#1,Quality:=USINT#2,Value:=LREAL#2.0,NowMs:=ULINT#5010,NominalDueMs:=ULINT#5000,SystemUtcMs:=ULINT#6000,Buffer:=Buffer);
    Policy(Buffer:=Buffer); phaseTicks:=0; Stage:=103;
103:
    Builder(GateOpen:=TRUE,NowMs:=Tick,UnixMs:=ULINT#7000,GatewayId:='test-gw',BootId:='test-boot',BatchIntervalMs:=UDINT#1,Buffer:=Buffer,Packets:=Packets,Sequence:=Sequence);
    phaseTicks:=phaseTicks+1;
    IF (Buffer.BatchOwners[1].State=2) OR (phaseTicks>500) THEN
        CheckIndex:=45; Check:=(Buffer.BatchOwners[1].Count=1) AND (FIND(Packets[1].Payload,CONCAT('"deviceId":',NG_Quote('changed"device')))>0) AND (FIND(Packets[1].Payload,NG_Quote('new"device'))=0);
        EndBatch(Slot:=UINT#1,Outcome:=USINT#2,Reason:=USINT#0,NowMs:=Tick,Buffer:=Buffer,Packets:=Packets);
        Stage:=104;
    END_IF;
104:
    Buffer.Configs[2]:=Buffer.Configs[1]; Buffer.ActiveSlot:=2;
    Buffer.Configs[2].Config.Devices[1].deviceId:='other"slot';
    Capture(PointIndex:=UINT#1,Kind:=USINT#1,Quality:=USINT#2,Value:=LREAL#3.0,NowMs:=ULINT#10010,NominalDueMs:=ULINT#10000,SystemUtcMs:=ULINT#11000,Buffer:=Buffer);
    Policy(Buffer:=Buffer); phaseTicks:=0; Stage:=105;
105:
    Builder(GateOpen:=TRUE,NowMs:=Tick,UnixMs:=ULINT#12000,GatewayId:='test-gw',BootId:='test-boot',BatchIntervalMs:=UDINT#1,Buffer:=Buffer,Packets:=Packets,Sequence:=Sequence);
    phaseTicks:=phaseTicks+1;
    IF (Buffer.BatchOwners[1].State=2) OR (phaseTicks>500) THEN
        CheckIndex:=46; Check:=(Buffer.BatchOwners[1].Count=1) AND (FIND(Packets[1].Payload,CONCAT('"deviceId":',NG_Quote('other"slot')))>0) AND (FIND(Packets[1].Payload,NG_Quote('changed"device'))=0);
        Stage:=106;
    END_IF;
106:
    Done:=TRUE;
END_CASE;
IF CheckIndex>0 THEN
    Checks[CheckIndex]:=Check;
    IF Check THEN Passed:=Passed+1; ELSE FailedChecks:=FailedChecks+1; END_IF;
END_IF;
END_PROGRAM

(* ---- platform_time_test.st ---- *)
PROGRAM Main
VAR
    LogicalClock : NG_PlatformTime;
    Permit : NG_TimePermit;
    WireTests : NG_TimeResponseTest;
    ClockDone : BOOL;
    Stage : UINT;
    Checks : ARRAY[1..40] OF BOOL;
    Passed : UINT;
    FailedChecks : UINT;
    Done : BOOL;
    Tick : ULINT := 100000;
    ResetClock : BOOL;
    Connected : BOOL := TRUE;
    Session : NG_Id := 'session-one';
    Submit : BOOL;
    Reply : BOOL;
    Heartbeat : BOOL;
    GetConfig : BOOL;
    RequestMono : ULINT;
    ServerT3 : ULINT;
    SystemDate : ULINT := 1000;
    SavedClockRevision : ULINT;
    SavedConnectionRevision : ULINT;
    SavedOutput : ULINT;
    Drift : LREAL := 50;
    i : UINT;
END_VAR
(* Offline assertion program. No gateway, socket, store, physical IO or RTC writes.
   Cold compilation is not execution; Done/Checks need a later authorized test runtime. *)
WireTests();
Done:=ClockDone AND WireTests.Done;
IF ClockDone THEN RETURN; END_IF;
ResetClock:=FALSE; Submit:=FALSE; Reply:=FALSE; Heartbeat:=FALSE; GetConfig:=FALSE;
CASE Stage OF
    0: ResetClock:=TRUE;
    1,3,5: Submit:=TRUE; RequestMono:=Tick;
    2,4,6: Tick:=Tick+20; Reply:=TRUE; ServerT3:=ULINT#1792000000000+Tick-100000-9;
    7: GetConfig:=TRUE;
    8: Heartbeat:=TRUE;
    9: GetConfig:=TRUE;
    10: SystemDate:=ULINT#9000000000000; Tick:=Tick+20;
    11: Connected:=FALSE; Tick:=Tick+20;
    12: Connected:=TRUE; Session:='session-two'; Tick:=Tick+20;
    13: Tick:=Tick+3600000;
    14: Tick:=Tick-1;
    15: ResetClock:=TRUE; Tick:=100000; Drift:=1000; Session:='recover-one';
    16,18,20,24,26,28,33,35,37,40,42,44,47,49,51,54,56,58: Submit:=TRUE; RequestMono:=Tick;
    17,19,21: Tick:=Tick+20; Reply:=TRUE; ServerT3:=ULINT#1792000000000+Tick-100000-9;
    22: SavedOutput:=LogicalClock.UtcMs; Connected:=FALSE; Tick:=Tick+172800000;
    23: Connected:=TRUE; Session:='recover-two';
    25,27,29: Tick:=Tick+20; Reply:=TRUE; ServerT3:=ULINT#1792000000000+Tick-100000-9-2170;
    30,60: Heartbeat:=TRUE;
    31,61: GetConfig:=TRUE;
    32,39: Tick:=Tick+330000;
    34,36,38: Tick:=Tick+20; Reply:=TRUE; ServerT3:=ULINT#1792000000000+Tick-100000-9-4340;
    41,43,45,48,50,52,55,57,59: Tick:=Tick+20; Reply:=TRUE; ServerT3:=ULINT#1792000000000+Tick-100000-9-90000;
    46: Tick:=Tick+10000;
    53: Tick:=Tick+120000;
END_CASE;
IF (Stage=37) OR (Stage=44) THEN SavedOutput:=LogicalClock.UtcMs; END_IF;
LogicalClock(Reset:=ResetClock,PlatformMode:=TRUE,Connected:=Connected,SessionId:=Session,NowMs:=Tick,SystemUtcMs:=SystemDate,
    TimeBasisRef:='site-hub-1',DriftBoundPpm:=Drift,DriftEvidence:='TEST_FIXTURE_ONLY',HistoryBasisRef:='',HistoryUtcLowerMs:=0,
    RequestSubmitted:=Submit,ResponseReady:=Reply,ResponseClientMonoMs:=RequestMono,ResponseReceivedMonoMs:=Tick,
    ServerReceivedMs:=ServerT3-2,ServerSentMs:=ServerT3,HeartbeatSubmitted:=Heartbeat,ConfigGetSubmitted:=GetConfig);
CASE Stage OF
0:
    Checks[1]:=LogicalClock.CaptureAllowed AND LogicalClock.AckApplyAllowed AND NOT LogicalClock.EnqueueAllowed AND NOT LogicalClock.ControlAllowed;
    Checks[2]:=LogicalClock.RequestWanted AND NOT LogicalClock.TimeValid;
1: Checks[3]:=LogicalClock.PendingRequest AND (LogicalClock.RequestClientMonoMs=Tick) AND (LogicalClock.Attempts=1);
2: Checks[4]:=NOT LogicalClock.TimeValid AND LogicalClock.RequestWanted;
6:
    Checks[5]:=LogicalClock.TimeValid AND LogicalClock.ControlAllowed AND NOT LogicalClock.SendAllowed;
    Checks[6]:=(LogicalClock.UtcMs=ULINT#1792000000060) AND (LogicalClock.UncertaintyMs=32);
    SavedClockRevision:=LogicalClock.ClockRevision; SavedConnectionRevision:=LogicalClock.ConnectionRevision;
7: Checks[7]:=NOT LogicalClock.SendAllowed;
8: Checks[8]:=NOT LogicalClock.SendAllowed;
9: Checks[9]:=LogicalClock.SendAllowed;
10: Checks[10]:=LogicalClock.TimeValid AND (LogicalClock.UtcMs=ULINT#1792000000080);
11: Checks[11]:=LogicalClock.TimeValid AND LogicalClock.EnqueueAllowed AND NOT LogicalClock.ControlAllowed AND NOT LogicalClock.SendAllowed;
12:
    Checks[12]:=LogicalClock.TimeValid AND NOT LogicalClock.ControlAllowed AND NOT LogicalClock.SendAllowed;
    Checks[13]:=(LogicalClock.ClockRevision=SavedClockRevision) AND (LogicalClock.ConnectionRevision>SavedConnectionRevision);
    Permit(Purpose:=USINT#4,TokenBootId:='boot-one',CurrentBootId:='boot-one',NowMs:=Tick,TokenMonoMs:=Tick,
        TokenClockRevision:=SavedClockRevision,TokenConnectionRevision:=SavedConnectionRevision,
        CurrentClockRevision:=LogicalClock.ClockRevision,CurrentConnectionRevision:=LogicalClock.ConnectionRevision,
        EnqueueAllowed:=TRUE,ControlAllowed:=TRUE,SendAllowed:=TRUE,AckApplyAllowed:=TRUE);
    Checks[14]:=NOT Permit.Allowed;
13:
    Checks[15]:=NOT LogicalClock.TimeValid AND NOT LogicalClock.EnqueueAllowed AND LogicalClock.CaptureAllowed AND LogicalClock.AckApplyAllowed;
    Checks[16]:=LogicalClock.State=4;
14:
    Checks[17]:=(LogicalClock.State=6) AND NOT LogicalClock.TimeValid;
    Permit(Purpose:=USINT#5,TokenBootId:='',CurrentBootId:='boot-one',NowMs:=Tick,TokenMonoMs:=0,
        TokenClockRevision:=0,TokenConnectionRevision:=0,CurrentClockRevision:=99,CurrentConnectionRevision:=99,
        EnqueueAllowed:=FALSE,ControlAllowed:=FALSE,SendAllowed:=FALSE,AckApplyAllowed:=TRUE);
    Checks[18]:=Permit.Allowed;
    Permit(Purpose:=USINT#2,TokenBootId:='old-boot',CurrentBootId:='boot-one',NowMs:=Tick,TokenMonoMs:=Tick,
        TokenClockRevision:=0,TokenConnectionRevision:=0,CurrentClockRevision:=0,CurrentConnectionRevision:=0,
        EnqueueAllowed:=TRUE,ControlAllowed:=TRUE,SendAllowed:=TRUE,AckApplyAllowed:=TRUE);
    Checks[19]:=NOT Permit.Allowed;
    Permit(Purpose:=USINT#2,TokenBootId:='boot-one',CurrentBootId:='boot-one',NowMs:=Tick,TokenMonoMs:=Tick-2000,
        TokenClockRevision:=0,TokenConnectionRevision:=0,CurrentClockRevision:=0,CurrentConnectionRevision:=0,
        EnqueueAllowed:=TRUE,ControlAllowed:=TRUE,SendAllowed:=TRUE,AckApplyAllowed:=TRUE);
    Checks[20]:=NOT Permit.Allowed;
    Permit(Purpose:=USINT#2,TokenBootId:='boot-one',CurrentBootId:='boot-one',NowMs:=Tick,TokenMonoMs:=Tick,
        TokenClockRevision:=0,TokenConnectionRevision:=0,CurrentClockRevision:=0,CurrentConnectionRevision:=0,
        EnqueueAllowed:=TRUE,ControlAllowed:=TRUE,SendAllowed:=TRUE,AckApplyAllowed:=TRUE);
    Checks[21]:=Permit.Allowed;
    LogicalClock(Reset:=TRUE,PlatformMode:=FALSE,Connected:=TRUE,SessionId:='compat',NowMs:=Tick,SystemUtcMs:=SystemDate,
        TimeBasisRef:='',DriftBoundPpm:=0,DriftEvidence:='',HistoryBasisRef:='',HistoryUtcLowerMs:=0,
        RequestSubmitted:=FALSE,ResponseReady:=FALSE,HeartbeatSubmitted:=FALSE,ConfigGetSubmitted:=FALSE);
    Checks[22]:=NOT LogicalClock.TimeValid AND LogicalClock.EnqueueAllowed AND NOT LogicalClock.RequestWanted;
    LogicalClock(Reset:=TRUE,PlatformMode:=TRUE,Connected:=TRUE,SessionId:='bad-drift',NowMs:=Tick,SystemUtcMs:=SystemDate,
        TimeBasisRef:='site-hub-1',DriftBoundPpm:=50,DriftEvidence:='',HistoryBasisRef:='',HistoryUtcLowerMs:=0);
    Checks[23]:=(LogicalClock.State=6) AND NOT LogicalClock.EnqueueAllowed;
    LogicalClock(Reset:=TRUE,PlatformMode:=TRUE,Connected:=TRUE,SessionId:='bad-basis',NowMs:=Tick,SystemUtcMs:=SystemDate,
        TimeBasisRef:='site-hub-1',DriftBoundPpm:=50,DriftEvidence:='TEST_FIXTURE_ONLY',HistoryBasisRef:='other-hub',HistoryUtcLowerMs:=1);
    Checks[24]:=(LogicalClock.State=6) AND NOT LogicalClock.EnqueueAllowed;
21: Checks[25]:=LogicalClock.TimeValid;
22: Checks[26]:=NOT LogicalClock.TimeValid AND (LogicalClock.State=4);
23: Checks[27]:=LogicalClock.RequestWanted;
29:
    Checks[28]:=LogicalClock.TimeValid;
    Checks[29]:=LogicalClock.State=2;
    Checks[30]:=LogicalClock.UtcMs>=SavedOutput;
    Checks[31]:=NOT LogicalClock.SendAllowed;
31: Checks[32]:=LogicalClock.SendAllowed;
38:
    Checks[33]:=LogicalClock.TimeValid AND (LogicalClock.UtcMs>=SavedOutput);
    Checks[34]:=(LogicalClock.State=2) AND (LogicalClock.UncertaintyMs<5000);
45: Checks[35]:=(LogicalClock.State=5) AND NOT LogicalClock.TimeValid;
46: Checks[36]:=LogicalClock.RequestWanted AND NOT LogicalClock.TimeValid;
52: Checks[37]:=(LogicalClock.State=4) AND NOT LogicalClock.TimeValid;
53: Checks[38]:=LogicalClock.RequestWanted;
59: Checks[39]:=LogicalClock.TimeValid AND (LogicalClock.UtcMs>=SavedOutput);
61:
    Checks[40]:=LogicalClock.TimeValid AND LogicalClock.SendAllowed AND (LogicalClock.State=2);
    Passed:=0; FailedChecks:=0;
    FOR i:=1 TO 40 DO IF Checks[i] THEN Passed:=Passed+1; ELSE FailedChecks:=FailedChecks+1; END_IF; END_FOR;
    ClockDone:=TRUE;
END_CASE;
Stage:=Stage+1;
END_PROGRAM
